Universal Robots URScript: FaiChun_9 Jan_11_2_t3.script

def Machining3():
  # Default parameters:
  global speed_ms = 0.05
  global speed_rads = 0.75
  global accel_mss = 3
  global accel_radss = 1.2
  global blend_radius_m = 0.0003

  # Add subprograms here
  # Start of main program
  # Program generated by RoboDK v5.6.8 for UR10e on 17/01/2025 15:25:47
  # Using nominal kinematics.
  blend_radius_m = 0.0003
  speed_ms = 0.05
  # set_reference(p[0.340000, 0.130000, 0.001500, 0.000000, 0.000000, 0.000000])
  set_tcp(p[0.000000, 0.000000, 0.252000, 0.000000, 0.000000, 0.000000])
  # Show Tool
  movej([0.835374, -1.505568, -2.356532, -0.850289, 1.570796, 2.406170],accel_radss,speed_rads,0,blend_radius_m)
  movel([0.835374, -1.553863, -2.383497, -0.775029, 1.570796, 2.406170],accel_mss,speed_ms,0,blend_radius_m)
  #SetTool1
  #M_RunCode6
  #SetRPM60000
  speed_ms = 0.05
  #M_RunCode3
  movel([0.835374, -1.574630, -2.393441, -0.744318, 1.570796, 2.406170],accel_mss,speed_ms,0,blend_radius_m)
  speed_ms = 0.003
  movel([0.835374, -1.579969, -2.395857, -0.736564, 1.570796, 2.406170],accel_mss,speed_ms,0,blend_radius_m)
  speed_ms = 0.015
  movel([0.633989, -1.489921, -2.480769, -0.741699, 1.570796, 2.204786],accel_mss,speed_ms,0,blend_radius_m)
  movel([0.864064, -1.190756, -2.677424, -0.844209, 1.570796, 2.434860],accel_mss,speed_ms,0,blend_radius_m)
  movel([1.072859, -1.363512, -2.578824, -0.770053, 1.570796, 2.643656],accel_mss,speed_ms,0,blend_radius_m)
  movel([0.835374, -1.579969, -2.395857, -0.736564, 1.570796, 2.406170],accel_mss,speed_ms,0,blend_radius_m)
  speed_ms = 0.003
  movel([0.835374, -1.574630, -2.393441, -0.744318, 1.570796, 2.406170],accel_mss,speed_ms,0,blend_radius_m)
  speed_ms = 0.05
  movel([0.835374, -1.553863, -2.383497, -0.775029, 1.570796, 2.406170],accel_mss,speed_ms,0,blend_radius_m)
  #M_RunCode9
  movel([0.837981, -1.545638, -2.391457, -0.775294, 1.570796, 2.408778],accel_mss,speed_ms,0,blend_radius_m)
  #M_RunCode3
  movel([0.837981, -1.566582, -2.401486, -0.744320, 1.570796, 2.408778],accel_mss,speed_ms,0,blend_radius_m)
  speed_ms = 0.003
  movel([0.837981, -1.571968, -2.403923, -0.736498, 1.570796, 2.408778],accel_mss,speed_ms,0,blend_radius_m)
  speed_ms = 0.012
  movel([0.835363, -1.570327, -2.405565, -0.736497, 1.570796, 2.406160],accel_mss,speed_ms,0,blend_radius_m)
  movel([0.832471, -1.573305, -2.402582, -0.736502, 1.570796, 2.403268],accel_mss,speed_ms,0,blend_radius_m)
  movel([0.828572, -1.570903, -2.404989, -0.736497, 1.570796, 2.399369],accel_mss,speed_ms,0,blend_radius_m)
  movel([0.831462, -1.567905, -2.407980, -0.736503, 1.570796, 2.402259],accel_mss,speed_ms,0,blend_radius_m)
  movel([0.830089, -1.567061, -2.408820, -0.736508, 1.570796, 2.400885],accel_mss,speed_ms,0,blend_radius_m)
  movel([0.827198, -1.570064, -2.405828, -0.736497, 1.570796, 2.397994],accel_mss,speed_ms,0,blend_radius_m)
  movel([0.823900, -1.568068, -2.407819, -0.736503, 1.570796, 2.394696],accel_mss,speed_ms,0,blend_radius_m)
  movel([0.823259, -1.567680, -2.408205, -0.736504, 1.570796, 2.394055],accel_mss,speed_ms,0,blend_radius_m)
  movel([0.827542, -1.563207, -2.412639, -0.736543, 1.570796, 2.398338],accel_mss,speed_ms,0,blend_radius_m)
  movel([0.830207, -1.564832, -2.411032, -0.736525, 1.570796, 2.401003],accel_mss,speed_ms,0,blend_radius_m)
  movel([0.831719, -1.563265, -2.412582, -0.736542, 1.570796, 2.402516],accel_mss,speed_ms,0,blend_radius_m)
  movel([0.827666, -1.560790, -2.415022, -0.736577, 1.570796, 2.398462],accel_mss,speed_ms,0,blend_radius_m)
  movel([0.821871, -1.566850, -2.409030, -0.736509, 1.570796, 2.392667],accel_mss,speed_ms,0,blend_radius_m)
  movel([0.821225, -1.566466, -2.409411, -0.736512, 1.570796, 2.392022],accel_mss,speed_ms,0,blend_radius_m)
  speed_ms = 0.02
  movel([0.744589, -1.526264, -2.448047, -0.738078, 1.570796, 2.315386],accel_mss,speed_ms,0,blend_radius_m)
  movel([0.657367, -1.492537, -2.478483, -0.741369, 1.570796, 2.228164],accel_mss,speed_ms,0,blend_radius_m)
  speed_ms = 0.012
  movel([0.662664, -1.485271, -2.484806, -0.742313, 1.570796, 2.233460],accel_mss,speed_ms,0,blend_radius_m)
  movel([0.657451, -1.483595, -2.486252, -0.742542, 1.570796, 2.228247],accel_mss,speed_ms,0,blend_radius_m)
  movel([0.656073, -1.485492, -2.484614, -0.742283, 1.570796, 2.226869],accel_mss,speed_ms,0,blend_radius_m)
  movel([0.659505, -1.486587, -2.483666, -0.742136, 1.570796, 2.230302],accel_mss,speed_ms,0,blend_radius_m)
  movel([0.655595, -1.491963, -2.478985, -0.741441, 1.570796, 2.226392],accel_mss,speed_ms,0,blend_radius_m)
  movel([0.654774, -1.491702, -2.479213, -0.741473, 1.570796, 2.225570],accel_mss,speed_ms,0,blend_radius_m)
  movel([0.650526, -1.490368, -2.480379, -0.741642, 1.570796, 2.221322],accel_mss,speed_ms,0,blend_radius_m)
  movel([0.653148, -1.486728, -2.483544, -0.742117, 1.570796, 2.223944],accel_mss,speed_ms,0,blend_radius_m)
  movel([0.651362, -1.486169, -2.484029, -0.742192, 1.570796, 2.222158],accel_mss,speed_ms,0,blend_radius_m)
  movel([0.648743, -1.489815, -2.480861, -0.741713, 1.570796, 2.219539],accel_mss,speed_ms,0,blend_radius_m)
  movel([0.643637, -1.488255, -2.482219, -0.741915, 1.570796, 2.214433],accel_mss,speed_ms,0,blend_radius_m)
  movel([0.646242, -1.484596, -2.485388, -0.742404, 1.570796, 2.217038],accel_mss,speed_ms,0,blend_radius_m)
  movel([0.642766, -1.483550, -2.486291, -0.742548, 1.570796, 2.213562],accel_mss,speed_ms,0,blend_radius_m)
  movel([0.646649, -1.478084, -2.490978, -0.743327, 1.570796, 2.217445],accel_mss,speed_ms,0,blend_radius_m)
  movel([0.650136, -1.479145, -2.490072, -0.743172, 1.570796, 2.220932],accel_mss,speed_ms,0,blend_radius_m)
  movel([0.651513, -1.477225, -2.491711, -0.743453, 1.570796, 2.222309],accel_mss,speed_ms,0,blend_radius_m)
  movel([0.648022, -1.476157, -2.492620, -0.743612, 1.570796, 2.218819],accel_mss,speed_ms,0,blend_radius_m)
  movel([0.651321, -1.471538, -2.496531, -0.744320, 1.570796, 2.222117],accel_mss,speed_ms,0,blend_radius_m)
  movel([0.651968, -1.470637, -2.497290, -0.744462, 1.570796, 2.222765],accel_mss,speed_ms,0,blend_radius_m)
  movel([0.657153, -1.472242, -2.495937, -0.744210, 1.570796, 2.227950],accel_mss,speed_ms,0,blend_radius_m)
  movel([0.654471, -1.475959, -2.492788, -0.743642, 1.570796, 2.225267],accel_mss,speed_ms,0,blend_radius_m)
  movel([0.656278, -1.476523, -2.492308, -0.743557, 1.570796, 2.227074],accel_mss,speed_ms,0,blend_radius_m)
  movel([0.660366, -1.470877, -2.497088, -0.744424, 1.570796, 2.231163],accel_mss,speed_ms,0,blend_radius_m)
  movel([0.653364, -1.468690, -2.498926, -0.744773, 1.570796, 2.224160],accel_mss,speed_ms,0,blend_radius_m)
  movel([0.735208, -1.358940, -2.581932, -0.771517, 1.570796, 2.306004],accel_mss,speed_ms,0,blend_radius_m)
  speed_ms = 0.02
  movel([0.838762, -1.228759, -2.658846, -0.824784, 1.570796, 2.409558],accel_mss,speed_ms,0,blend_radius_m)
  movel([0.839821, -1.227466, -2.659505, -0.825418, 1.570796, 2.410617],accel_mss,speed_ms,0,blend_radius_m)
  speed_ms = 0.012
  movel([0.847664, -1.231537, -2.657424, -0.823428, 1.570796, 2.418460],accel_mss,speed_ms,0,blend_radius_m)
  movel([0.854413, -1.223391, -2.661569, -0.827429, 1.570796, 2.425209],accel_mss,speed_ms,0,blend_radius_m)
  movel([0.852387, -1.222304, -2.662116, -0.827969, 1.570796, 2.423183],accel_mss,speed_ms,0,blend_radius_m)
  movel([0.847934, -1.227691, -2.659391, -0.825307, 1.570796, 2.418730],accel_mss,speed_ms,0,blend_radius_m)
  movel([0.842121, -1.224661, -2.660928, -0.826800, 1.570796, 2.412917],accel_mss,speed_ms,0,blend_radius_m)
  movel([0.843184, -1.223362, -2.661584, -0.827444, 1.570796, 2.413980],accel_mss,speed_ms,0,blend_radius_m)
  movel([0.848718, -1.216604, -2.664964, -0.830821, 1.570796, 2.419515],accel_mss,speed_ms,0,blend_radius_m)
  movel([0.852657, -1.218688, -2.663927, -0.829774, 1.570796, 2.423453],accel_mss,speed_ms,0,blend_radius_m)
  movel([0.854994, -1.215856, -2.665335, -0.831197, 1.570796, 2.425791],accel_mss,speed_ms,0,blend_radius_m)
  movel([0.851054, -1.213757, -2.666373, -0.832259, 1.570796, 2.421850],accel_mss,speed_ms,0,blend_radius_m)
  movel([0.857788, -1.205562, -2.670377, -0.836450, 1.570796, 2.428584],accel_mss,speed_ms,0,blend_radius_m)
  movel([0.861735, -1.207706, -2.669337, -0.835346, 1.570796, 2.432532],accel_mss,speed_ms,0,blend_radius_m)
  movel([0.866344, -1.202146, -2.672025, -0.838219, 1.570796, 2.437140],accel_mss,speed_ms,0,blend_radius_m)
  movel([0.872146, -1.205404, -2.670454, -0.836531, 1.570796, 2.442943],accel_mss,speed_ms,0,blend_radius_m)
  movel([0.867532, -1.210918, -2.667769, -0.833702, 1.570796, 2.438328],accel_mss,speed_ms,0,blend_radius_m)
  movel([0.869549, -1.212054, -2.667212, -0.833124, 1.570796, 2.440345],accel_mss,speed_ms,0,blend_radius_m)
  movel([0.874165, -1.206556, -2.669896, -0.835937, 1.570796, 2.444961],accel_mss,speed_ms,0,blend_radius_m)
  movel([0.879884, -1.209871, -2.668281, -0.834237, 1.570796, 2.450680],accel_mss,speed_ms,0,blend_radius_m)
  movel([0.873058, -1.217928, -2.664306, -0.830155, 1.570796, 2.443854],accel_mss,speed_ms,0,blend_radius_m)
  movel([0.869206, -1.215731, -2.665397, -0.831261, 1.570796, 2.440003],accel_mss,speed_ms,0,blend_radius_m)
  movel([0.866837, -1.218550, -2.663996, -0.829843, 1.570796, 2.437634],accel_mss,speed_ms,0,blend_radius_m)
  movel([0.872676, -1.221871, -2.662334, -0.828184, 1.570796, 2.443472],accel_mss,speed_ms,0,blend_radius_m)
  movel([0.881873, -1.211042, -2.667708, -0.833639, 1.570796, 2.452670],accel_mss,speed_ms,0,blend_radius_m)
  movel([0.975719, -1.277693, -2.632456, -0.802240, 1.570796, 2.546515],accel_mss,speed_ms,0,blend_radius_m)
  speed_ms = 0.02
  movel([1.052001, -1.350806, -2.587390, -0.774193, 1.570796, 2.622798],accel_mss,speed_ms,0,blend_radius_m)
  movel([1.043190, -1.358370, -2.582317, -0.771702, 1.570796, 2.613987],accel_mss,speed_ms,0,blend_radius_m)
  speed_ms = 0.012
  movel([1.047039, -1.362473, -2.579533, -0.770383, 1.570796, 2.617836],accel_mss,speed_ms,0,blend_radius_m)
  movel([1.049307, -1.360540, -2.580848, -0.771002, 1.570796, 2.620103],accel_mss,speed_ms,0,blend_radius_m)
  movel([1.046783, -1.357825, -2.582685, -0.771878, 1.570796, 2.617579],accel_mss,speed_ms,0,blend_radius_m)
  movel([1.053311, -1.352246, -2.586430, -0.773713, 1.570796, 2.624108],accel_mss,speed_ms,0,blend_radius_m)
  movel([1.053918, -1.352909, -2.585988, -0.773493, 1.570796, 2.624714],accel_mss,speed_ms,0,blend_radius_m)
  movel([1.057025, -1.356325, -2.583697, -0.772367, 1.570796, 2.627821],accel_mss,speed_ms,0,blend_radius_m)
  movel([1.052623, -1.360057, -2.581176, -0.771157, 1.570796, 2.623420],accel_mss,speed_ms,0,blend_radius_m)
  movel([1.053917, -1.361475, -2.580212, -0.770702, 1.570796, 2.624713],accel_mss,speed_ms,0,blend_radius_m)
  movel([1.058318, -1.357758, -2.582731, -0.771900, 1.570796, 2.629115],accel_mss,speed_ms,0,blend_radius_m)
  movel([1.061975, -1.361842, -2.579962, -0.770584, 1.570796, 2.632771],accel_mss,speed_ms,0,blend_radius_m)
  movel([1.057587, -1.365521, -2.577449, -0.769419, 1.570796, 2.628383],accel_mss,speed_ms,0,blend_radius_m)
  movel([1.060041, -1.368254, -2.575569, -0.768566, 1.570796, 2.630837],accel_mss,speed_ms,0,blend_radius_m)
  movel([1.053613, -1.373635, -2.571837, -0.766917, 1.570796, 2.624409],accel_mss,speed_ms,0,blend_radius_m)
  movel([1.051147, -1.370941, -2.573711, -0.767737, 1.570796, 2.621943],accel_mss,speed_ms,0,blend_radius_m)
  movel([1.048905, -1.372833, -2.572396, -0.767160, 1.570796, 2.619702],accel_mss,speed_ms,0,blend_radius_m)
  movel([1.051373, -1.375516, -2.570523, -0.766350, 1.570796, 2.622169],accel_mss,speed_ms,0,blend_radius_m)
  movel([1.046058, -1.379991, -2.567376, -0.765022, 1.570796, 2.616855],accel_mss,speed_ms,0,blend_radius_m)
  movel([1.045032, -1.380857, -2.566764, -0.764768, 1.570796, 2.615828],accel_mss,speed_ms,0,blend_radius_m)
  movel([1.041351, -1.376942, -2.569524, -0.765924, 1.570796, 2.612147],accel_mss,speed_ms,0,blend_radius_m)
  movel([1.045637, -1.373301, -2.572070, -0.767018, 1.570796, 2.616433],accel_mss,speed_ms,0,blend_radius_m)
  movel([1.044340, -1.371916, -2.573034, -0.767439, 1.570796, 2.615136],accel_mss,speed_ms,0,blend_radius_m)
  movel([1.037833, -1.377462, -2.569158, -0.765769, 1.570796, 2.608629],accel_mss,speed_ms,0,blend_radius_m)
  movel([1.042823, -1.382724, -2.565440, -0.764225, 1.570796, 2.613619],accel_mss,speed_ms,0,blend_radius_m)
  speed_ms = 0.02
  movel([0.937722, -1.475331, -2.493322, -0.743736, 1.570796, 2.508518],accel_mss,speed_ms,0,blend_radius_m)
  movel([0.849748, -1.560014, -2.415785, -0.736589, 1.570796, 2.420545],accel_mss,speed_ms,0,blend_radius_m)
  speed_ms = 0.012
  movel([0.844480, -1.556645, -2.419087, -0.736656, 1.570796, 2.415277],accel_mss,speed_ms,0,blend_radius_m)
  movel([0.839983, -1.561236, -2.414583, -0.736570, 1.570796, 2.410779],accel_mss,speed_ms,0,blend_radius_m)
  movel([0.841353, -1.562100, -2.413732, -0.736557, 1.570796, 2.412149],accel_mss,speed_ms,0,blend_radius_m)
  movel([0.844308, -1.559087, -2.416696, -0.736606, 1.570796, 2.415104],accel_mss,speed_ms,0,blend_radius_m)
  movel([0.848197, -1.561574, -2.414251, -0.736565, 1.570796, 2.418993],accel_mss,speed_ms,0,blend_radius_m)
  movel([0.847483, -1.562295, -2.413539, -0.736554, 1.570796, 2.418279],accel_mss,speed_ms,0,blend_radius_m)
  movel([0.843823, -1.566008, -2.409866, -0.736515, 1.570796, 2.414620],accel_mss,speed_ms,0,blend_radius_m)
  movel([0.841203, -1.564344, -2.411515, -0.736530, 1.570796, 2.411999],accel_mss,speed_ms,0,blend_radius_m)
  movel([0.839681, -1.565899, -2.409974, -0.736516, 1.570796, 2.410477],accel_mss,speed_ms,0,blend_radius_m)
  movel([0.842302, -1.567558, -2.408326, -0.736505, 1.570796, 2.413098],accel_mss,speed_ms,0,blend_radius_m)
  movel([0.837981, -1.571968, -2.403923, -0.736498, 1.570796, 2.408778],accel_mss,speed_ms,0,blend_radius_m)
  speed_ms = 0.003
  movel([0.837981, -1.566582, -2.401486, -0.744320, 1.570796, 2.408778],accel_mss,speed_ms,0,blend_radius_m)
  speed_ms = 0.05
  movel([0.837981, -1.545638, -2.391457, -0.775294, 1.570796, 2.408778],accel_mss,speed_ms,0,blend_radius_m)
  #M_RunCode9
  movel([0.855198, -1.260338, -2.606468, -0.845583, 1.570796, 2.425994],accel_mss,speed_ms,0,blend_radius_m)
  #M_RunCode3
  # num 0 inside
  movel([0.855198, -1.286686, -2.619958, -0.805745, 1.570796, 2.425994],accel_mss,speed_ms,0,blend_radius_m)
  speed_ms = 0.003
  movel([0.855198, -1.293571, -2.623261, -0.795557, 1.570796, 2.425994],accel_mss,speed_ms,0,blend_radius_m)
  speed_ms = 0.015
  movel([0.846910, -1.296288, -2.621656, -0.794445, 1.570796, 2.417706],accel_mss,speed_ms,0,blend_radius_m)
  movel([0.841111, -1.297727, -2.620801, -0.793860, 1.570796, 2.411907],accel_mss,speed_ms,0,blend_radius_m)
  movel([0.839123, -1.297920, -2.620687, -0.793782, 1.570796, 2.409919],accel_mss,speed_ms,0,blend_radius_m)
  movel([0.837725, -1.297694, -2.620821, -0.793874, 1.570796, 2.408522],accel_mss,speed_ms,0,blend_radius_m)
  movel([0.836916, -1.297054, -2.621202, -0.794134, 1.570796, 2.407712],accel_mss,speed_ms,0,blend_radius_m)
  movel([0.836696, -1.295992, -2.621831, -0.794566, 1.570796, 2.407493],accel_mss,speed_ms,0,blend_radius_m)
  movel([0.837055, -1.294718, -2.622585, -0.795086, 1.570796, 2.407851],accel_mss,speed_ms,0,blend_radius_m)
  movel([0.837982, -1.293440, -2.623338, -0.795611, 1.570796, 2.408779],accel_mss,speed_ms,0,blend_radius_m)
  movel([0.839480, -1.292159, -2.624092, -0.796138, 1.570796, 2.410276],accel_mss,speed_ms,0,blend_radius_m)
  movel([0.841550, -1.290874, -2.624846, -0.796670, 1.570796, 2.412346],accel_mss,speed_ms,0,blend_radius_m)
  movel([0.847491, -1.288081, -2.626476, -0.797832, 1.570796, 2.418287],accel_mss,speed_ms,0,blend_radius_m)
  movel([0.855893, -1.284860, -2.628345, -0.799184, 1.570796, 2.426689],accel_mss,speed_ms,0,blend_radius_m)
  movel([0.864286, -1.282119, -2.629925, -0.800345, 1.570796, 2.435082],accel_mss,speed_ms,0,blend_radius_m)
  movel([0.870165, -1.280730, -2.630722, -0.800937, 1.570796, 2.440961],accel_mss,speed_ms,0,blend_radius_m)
  movel([0.872167, -1.280581, -2.630807, -0.801001, 1.570796, 2.442964],accel_mss,speed_ms,0,blend_radius_m)
  movel([0.873560, -1.280853, -2.630651, -0.800885, 1.570796, 2.444356],accel_mss,speed_ms,0,blend_radius_m)
  movel([0.874341, -1.281545, -2.630255, -0.800590, 1.570796, 2.445137],accel_mss,speed_ms,0,blend_radius_m)
  movel([0.874513, -1.282655, -2.629617, -0.800118, 1.570796, 2.445309],accel_mss,speed_ms,0,blend_radius_m)
  movel([0.874099, -1.283962, -2.628863, -0.799563, 1.570796, 2.444895],accel_mss,speed_ms,0,blend_radius_m)
  movel([0.873124, -1.285249, -2.628120, -0.799020, 1.570796, 2.443921],accel_mss,speed_ms,0,blend_radius_m)
  movel([0.871587, -1.286518, -2.627385, -0.798486, 1.570796, 2.442383],accel_mss,speed_ms,0,blend_radius_m)
  movel([0.869494, -1.287766, -2.626660, -0.797963, 1.570796, 2.440290],accel_mss,speed_ms,0,blend_radius_m)
  movel([0.863543, -1.290454, -2.625092, -0.796844, 1.570796, 2.434339],accel_mss,speed_ms,0,blend_radius_m)
  movel([0.855198, -1.293571, -2.623261, -0.795557, 1.570796, 2.425994],accel_mss,speed_ms,0,blend_radius_m)
  speed_ms = 0.003
  movel([0.855198, -1.286686, -2.619958, -0.805745, 1.570796, 2.425994],accel_mss,speed_ms,0,blend_radius_m)
  speed_ms = 0.05
  movel([0.855198, -1.260338, -2.606468, -0.845583, 1.570796, 2.425994],accel_mss,speed_ms,0,blend_radius_m)
  #M_RunCode9
  movel([0.854459, -1.269799, -2.601095, -0.841495, 1.570796, 2.425256],accel_mss,speed_ms,0,blend_radius_m)
  #M_RunCode3
  #num 0 outside
  movel([0.854459, -1.296016, -2.614460, -0.801913, 1.570796, 2.425256],accel_mss,speed_ms,0,blend_radius_m)
  speed_ms = 0.003
  movel([0.854459, -1.302862, -2.617732, -0.791795, 1.570796, 2.425256],accel_mss,speed_ms,0,blend_radius_m)
  speed_ms = 0.015
  movel([0.851475, -1.303789, -2.617174, -0.791426, 1.570796, 2.422272],accel_mss,speed_ms,0,blend_radius_m)
  movel([0.848730, -1.304421, -2.616793, -0.791175, 1.570796, 2.419526],accel_mss,speed_ms,0,blend_radius_m)
  movel([0.846217, -1.304761, -2.616588, -0.791040, 1.570796, 2.417014],accel_mss,speed_ms,0,blend_radius_m)
  movel([0.843939, -1.304807, -2.616560, -0.791022, 1.570796, 2.414735],accel_mss,speed_ms,0,blend_radius_m)
  movel([0.841916, -1.304581, -2.616697, -0.791111, 1.570796, 2.412713],accel_mss,speed_ms,0,blend_radius_m)
  movel([0.840172, -1.304105, -2.616984, -0.791300, 1.570796, 2.410968],accel_mss,speed_ms,0,blend_radius_m)
  movel([0.838702, -1.303380, -2.617420, -0.791589, 1.570796, 2.409498],accel_mss,speed_ms,0,blend_radius_m)
  movel([0.837514, -1.302400, -2.618010, -0.791979, 1.570796, 2.408310],accel_mss,speed_ms,0,blend_radius_m)
  movel([0.836610, -1.301192, -2.618734, -0.792463, 1.570796, 2.407406],accel_mss,speed_ms,0,blend_radius_m)
  movel([0.835994, -1.299790, -2.619572, -0.793026, 1.570796, 2.406790],accel_mss,speed_ms,0,blend_radius_m)
  movel([0.835668, -1.298186, -2.620529, -0.793674, 1.570796, 2.406464],accel_mss,speed_ms,0,blend_radius_m)
  movel([0.835631, -1.296383, -2.621599, -0.794407, 1.570796, 2.406427],accel_mss,speed_ms,0,blend_radius_m)
  movel([0.835884, -1.294466, -2.622733, -0.795190, 1.570796, 2.406680],accel_mss,speed_ms,0,blend_radius_m)
  movel([0.836421, -1.292534, -2.623871, -0.795983, 1.570796, 2.407217],accel_mss,speed_ms,0,blend_radius_m)
  movel([0.837240, -1.290586, -2.625014, -0.796789, 1.570796, 2.408036],accel_mss,speed_ms,0,blend_radius_m)
  movel([0.838350, -1.288617, -2.626164, -0.797608, 1.570796, 2.409146],accel_mss,speed_ms,0,blend_radius_m)
  movel([0.839739, -1.286668, -2.627298, -0.798423, 1.570796, 2.410536],accel_mss,speed_ms,0,blend_radius_m)
  movel([0.841401, -1.284772, -2.628396, -0.799221, 1.570796, 2.412197],accel_mss,speed_ms,0,blend_radius_m)
  movel([0.843338, -1.282931, -2.629458, -0.800000, 1.570796, 2.414134],accel_mss,speed_ms,0,blend_radius_m)
  movel([0.845550, -1.281147, -2.630483, -0.800759, 1.570796, 2.416347],accel_mss,speed_ms,0,blend_radius_m)
  movel([0.848009, -1.279462, -2.631447, -0.801480, 1.570796, 2.418805],accel_mss,speed_ms,0,blend_radius_m)
  movel([0.850682, -1.277926, -2.632323, -0.802140, 1.570796, 2.421478],accel_mss,speed_ms,0,blend_radius_m)
  movel([0.853567, -1.276542, -2.633110, -0.802737, 1.570796, 2.424364],accel_mss,speed_ms,0,blend_radius_m)
  movel([0.856663, -1.275312, -2.633807, -0.803270, 1.570796, 2.427459],accel_mss,speed_ms,0,blend_radius_m)
  movel([0.859747, -1.274318, -2.634369, -0.803702, 1.570796, 2.430544],accel_mss,speed_ms,0,blend_radius_m)
  movel([0.862585, -1.273645, -2.634749, -0.803995, 1.570796, 2.433381],accel_mss,speed_ms,0,blend_radius_m)
  movel([0.865178, -1.273292, -2.634948, -0.804149, 1.570796, 2.435974],accel_mss,speed_ms,0,blend_radius_m)
  movel([0.867519, -1.273260, -2.634966, -0.804163, 1.570796, 2.438315],accel_mss,speed_ms,0,blend_radius_m)
  movel([0.869584, -1.273524, -2.634817, -0.804048, 1.570796, 2.440380],accel_mss,speed_ms,0,blend_radius_m)
  movel([0.871341, -1.274060, -2.634515, -0.803814, 1.570796, 2.442138],accel_mss,speed_ms,0,blend_radius_m)
  movel([0.872797, -1.274863, -2.634061, -0.803465, 1.570796, 2.443593],accel_mss,speed_ms,0,blend_radius_m)
  movel([0.873946, -1.275936, -2.633454, -0.803000, 1.570796, 2.444743],accel_mss,speed_ms,0,blend_radius_m)
  movel([0.874790, -1.277237, -2.632715, -0.802437, 1.570796, 2.445586],accel_mss,speed_ms,0,blend_radius_m)
  movel([0.875334, -1.278736, -2.631862, -0.801792, 1.570796, 2.446131],accel_mss,speed_ms,0,blend_radius_m)
  movel([0.875580, -1.280428, -2.630895, -0.801066, 1.570796, 2.446377],accel_mss,speed_ms,0,blend_radius_m)
  movel([0.875527, -1.282310, -2.629815, -0.800264, 1.570796, 2.446323],accel_mss,speed_ms,0,blend_radius_m)
  movel([0.875187, -1.284285, -2.628677, -0.799427, 1.570796, 2.445983],accel_mss,speed_ms,0,blend_radius_m)
  movel([0.874574, -1.286253, -2.627538, -0.798598, 1.570796, 2.445370],accel_mss,speed_ms,0,blend_radius_m)
  movel([0.873688, -1.288215, -2.626398, -0.797776, 1.570796, 2.444484],accel_mss,speed_ms,0,blend_radius_m)
  movel([0.872531, -1.290171, -2.625257, -0.796961, 1.570796, 2.443327],accel_mss,speed_ms,0,blend_radius_m)
  movel([0.871111, -1.292085, -2.624135, -0.796169, 1.570796, 2.441907],accel_mss,speed_ms,0,blend_radius_m)
  movel([0.869432, -1.293928, -2.623051, -0.795410, 1.570796, 2.440228],accel_mss,speed_ms,0,blend_radius_m)
  movel([0.867493, -1.295700, -2.622004, -0.794685, 1.570796, 2.438289],accel_mss,speed_ms,0,blend_radius_m)
  movel([0.865298, -1.297400, -2.620996, -0.793993, 1.570796, 2.436095],accel_mss,speed_ms,0,blend_radius_m)
  movel([0.862881, -1.298989, -2.620050, -0.793350, 1.570796, 2.433677],accel_mss,speed_ms,0,blend_radius_m)
  movel([0.860267, -1.300428, -2.619191, -0.792770, 1.570796, 2.431063],accel_mss,speed_ms,0,blend_radius_m)
  movel([0.857460, -1.301718, -2.618419, -0.792252, 1.570796, 2.428257],accel_mss,speed_ms,0,blend_radius_m)
  movel([0.854459, -1.302862, -2.617732, -0.791795, 1.570796, 2.425256],accel_mss,speed_ms,0,blend_radius_m)
  speed_ms = 0.003
  movel([0.854459, -1.296016, -2.614460, -0.801913, 1.570796, 2.425256],accel_mss,speed_ms,0,blend_radius_m)
  speed_ms = 0.05
  movel([0.854459, -1.269799, -2.601095, -0.841495, 1.570796, 2.425256],accel_mss,speed_ms,0,blend_radius_m)
  #M_RunCode9
  movel([0.848212, -1.241330, -2.616943, -0.854116, 1.570796, 2.419008],accel_mss,speed_ms,0,blend_radius_m)
  #M_RunCode3
  # num 2
  movel([0.848212, -1.267925, -2.630682, -0.813782, 1.570796, 2.419008],accel_mss,speed_ms,0,blend_radius_m)
  speed_ms = 0.003
  movel([0.848212, -1.274884, -2.634049, -0.803455, 1.570796, 2.419008],accel_mss,speed_ms,0,blend_radius_m)
  speed_ms = 0.02
  movel([0.837317, -1.278925, -2.631754, -0.801710, 1.570796, 2.408113],accel_mss,speed_ms,0,blend_radius_m)
  movel([0.839074, -1.249773, -2.647865, -0.814751, 1.570796, 2.409870],accel_mss,speed_ms,0,blend_radius_m)
  movel([0.840196, -1.249335, -2.648099, -0.814955, 1.570796, 2.410992],accel_mss,speed_ms,0,blend_radius_m)
  movel([0.843034, -1.248564, -2.648511, -0.815314, 1.570796, 2.413831],accel_mss,speed_ms,0,blend_radius_m)
  movel([0.845771, -1.248506, -2.648542, -0.815341, 1.570796, 2.416567],accel_mss,speed_ms,0,blend_radius_m)
  movel([0.848339, -1.248990, -2.648284, -0.815116, 1.570796, 2.419136],accel_mss,speed_ms,0,blend_radius_m)
  movel([0.850670, -1.249839, -2.647829, -0.814720, 1.570796, 2.421467],accel_mss,speed_ms,0,blend_radius_m)
  movel([0.856325, -1.252900, -2.646186, -0.813303, 1.570796, 2.427121],accel_mss,speed_ms,0,blend_radius_m)
  movel([0.861461, -1.255841, -2.644597, -0.811951, 1.570796, 2.432257],accel_mss,speed_ms,0,blend_radius_m)
  movel([0.863580, -1.256692, -2.644135, -0.811562, 1.570796, 2.434377],accel_mss,speed_ms,0,blend_radius_m)
  movel([0.865859, -1.257203, -2.643857, -0.811329, 1.570796, 2.436655],accel_mss,speed_ms,0,blend_radius_m)
  movel([0.868233, -1.257243, -2.643835, -0.811311, 1.570796, 2.439030],accel_mss,speed_ms,0,blend_radius_m)
  movel([0.870648, -1.256675, -2.644144, -0.811570, 1.570796, 2.441444],accel_mss,speed_ms,0,blend_radius_m)
  movel([0.873569, -1.255238, -2.644923, -0.812228, 1.570796, 2.444365],accel_mss,speed_ms,0,blend_radius_m)
  movel([0.874767, -1.254321, -2.645420, -0.812649, 1.570796, 2.445563],accel_mss,speed_ms,0,blend_radius_m)
  movel([0.875791, -1.253271, -2.645986, -0.813132, 1.570796, 2.446587],accel_mss,speed_ms,0,blend_radius_m)
  movel([0.877258, -1.251040, -2.647186, -0.814163, 1.570796, 2.448054],accel_mss,speed_ms,0,blend_radius_m)
  movel([0.877898, -1.248826, -2.648371, -0.815192, 1.570796, 2.448694],accel_mss,speed_ms,0,blend_radius_m)
  movel([0.877875, -1.247491, -2.649083, -0.815815, 1.570796, 2.448671],accel_mss,speed_ms,0,blend_radius_m)
  movel([0.877482, -1.246635, -2.649538, -0.816216, 1.570796, 2.448278],accel_mss,speed_ms,0,blend_radius_m)
  movel([0.876798, -1.246264, -2.649735, -0.816390, 1.570796, 2.447594],accel_mss,speed_ms,0,blend_radius_m)
  movel([0.875913, -1.246377, -2.649675, -0.816337, 1.570796, 2.446709],accel_mss,speed_ms,0,blend_radius_m)
  movel([0.874526, -1.247366, -2.649149, -0.815874, 1.570796, 2.445322],accel_mss,speed_ms,0,blend_radius_m)
  movel([0.873202, -1.248420, -2.648588, -0.815381, 1.570796, 2.443999],accel_mss,speed_ms,0,blend_radius_m)
  movel([0.871495, -1.249252, -2.648143, -0.814993, 1.570796, 2.442292],accel_mss,speed_ms,0,blend_radius_m)
  movel([0.869538, -1.249620, -2.647947, -0.814822, 1.570796, 2.440334],accel_mss,speed_ms,0,blend_radius_m)
  movel([0.868153, -1.249104, -2.648222, -0.815062, 1.570796, 2.438950],accel_mss,speed_ms,0,blend_radius_m)
  movel([0.867374, -1.247895, -2.648867, -0.815626, 1.570796, 2.438171],accel_mss,speed_ms,0,blend_radius_m)
  movel([0.867234, -1.246189, -2.649775, -0.816425, 1.570796, 2.438030],accel_mss,speed_ms,0,blend_radius_m)
  movel([0.867710, -1.244254, -2.650799, -0.817336, 1.570796, 2.438506],accel_mss,speed_ms,0,blend_radius_m)
  movel([0.868781, -1.242353, -2.651802, -0.818234, 1.570796, 2.439578],accel_mss,speed_ms,0,blend_radius_m)
  movel([0.870379, -1.240727, -2.652656, -0.819006, 1.570796, 2.441175],accel_mss,speed_ms,0,blend_radius_m)
  movel([0.872426, -1.239628, -2.653231, -0.819530, 1.570796, 2.443223],accel_mss,speed_ms,0,blend_radius_m)
  movel([0.874179, -1.239185, -2.653463, -0.819741, 1.570796, 2.444975],accel_mss,speed_ms,0,blend_radius_m)
  movel([0.875671, -1.239239, -2.653435, -0.819716, 1.570796, 2.446467],accel_mss,speed_ms,0,blend_radius_m)
  movel([0.876905, -1.239788, -2.653148, -0.819454, 1.570796, 2.447701],accel_mss,speed_ms,0,blend_radius_m)
  movel([0.877875, -1.240835, -2.652599, -0.818955, 1.570796, 2.448672],accel_mss,speed_ms,0,blend_radius_m)
  movel([0.878573, -1.242283, -2.651839, -0.818268, 1.570796, 2.449370],accel_mss,speed_ms,0,blend_radius_m)
  movel([0.878998, -1.244031, -2.650917, -0.817441, 1.570796, 2.449794],accel_mss,speed_ms,0,blend_radius_m)
  movel([0.879021, -1.248427, -2.648584, -0.815378, 1.570796, 2.449817],accel_mss,speed_ms,0,blend_radius_m)
  movel([0.878543, -1.251428, -2.646978, -0.813983, 1.570796, 2.449340],accel_mss,speed_ms,0,blend_radius_m)
  movel([0.877746, -1.254377, -2.645389, -0.812623, 1.570796, 2.448542],accel_mss,speed_ms,0,blend_radius_m)
  movel([0.876632, -1.257271, -2.643820, -0.811298, 1.570796, 2.447428],accel_mss,speed_ms,0,blend_radius_m)
  movel([0.875201, -1.260113, -2.642269, -0.810007, 1.570796, 2.445997],accel_mss,speed_ms,0,blend_radius_m)
  movel([0.873417, -1.262713, -2.640842, -0.808835, 1.570796, 2.444214],accel_mss,speed_ms,0,blend_radius_m)
  movel([0.871230, -1.264887, -2.639642, -0.807860, 1.570796, 2.442027],accel_mss,speed_ms,0,blend_radius_m)
  movel([0.868642, -1.266641, -2.638669, -0.807078, 1.570796, 2.439438],accel_mss,speed_ms,0,blend_radius_m)
  movel([0.865652, -1.267984, -2.637922, -0.806483, 1.570796, 2.436448],accel_mss,speed_ms,0,blend_radius_m)
  movel([0.862952, -1.268698, -2.637524, -0.806167, 1.570796, 2.433748],accel_mss,speed_ms,0,blend_radius_m)
  movel([0.860488, -1.268833, -2.637449, -0.806107, 1.570796, 2.431284],accel_mss,speed_ms,0,blend_radius_m)
  movel([0.858259, -1.268518, -2.637624, -0.806246, 1.570796, 2.429055],accel_mss,speed_ms,0,blend_radius_m)
  movel([0.856267, -1.267886, -2.637977, -0.806526, 1.570796, 2.427063],accel_mss,speed_ms,0,blend_radius_m)
  movel([0.851897, -1.265592, -2.639251, -0.807546, 1.570796, 2.422694],accel_mss,speed_ms,0,blend_radius_m)
  movel([0.847719, -1.263475, -2.640421, -0.808492, 1.570796, 2.418515],accel_mss,speed_ms,0,blend_radius_m)
  movel([0.845888, -1.262909, -2.640734, -0.808746, 1.570796, 2.416685],accel_mss,speed_ms,0,blend_radius_m)
  movel([0.843868, -1.262640, -2.640882, -0.808867, 1.570796, 2.414664],accel_mss,speed_ms,0,blend_radius_m)
  movel([0.841671, -1.262784, -2.640803, -0.808803, 1.570796, 2.412467],accel_mss,speed_ms,0,blend_radius_m)
  movel([0.839325, -1.263447, -2.640437, -0.808505, 1.570796, 2.410122],accel_mss,speed_ms,0,blend_radius_m)
  movel([0.839258, -1.264541, -2.639833, -0.808015, 1.570796, 2.410054],accel_mss,speed_ms,0,blend_radius_m)
  movel([0.839240, -1.267497, -2.638194, -0.806699, 1.570796, 2.410037],accel_mss,speed_ms,0,blend_radius_m)
  movel([0.839588, -1.269943, -2.636829, -0.805617, 1.570796, 2.410384],accel_mss,speed_ms,0,blend_radius_m)
  movel([0.840292, -1.271889, -2.635738, -0.804762, 1.570796, 2.411089],accel_mss,speed_ms,0,blend_radius_m)
  movel([0.841357, -1.273337, -2.634923, -0.804129, 1.570796, 2.412154],accel_mss,speed_ms,0,blend_radius_m)
  movel([0.842716, -1.274334, -2.634360, -0.803695, 1.570796, 2.413512],accel_mss,speed_ms,0,blend_radius_m)
  movel([0.844310, -1.274923, -2.634027, -0.803439, 1.570796, 2.415107],accel_mss,speed_ms,0,blend_radius_m)
  movel([0.846140, -1.275106, -2.633924, -0.803359, 1.570796, 2.416937],accel_mss,speed_ms,0,blend_radius_m)
  movel([0.848212, -1.274884, -2.634049, -0.803455, 1.570796, 2.419008],accel_mss,speed_ms,0,blend_radius_m)
  speed_ms = 0.003
  movel([0.848212, -1.267925, -2.630682, -0.813782, 1.570796, 2.419008],accel_mss,speed_ms,0,blend_radius_m)
  speed_ms = 0.05
  movel([0.848212, -1.241330, -2.616943, -0.854116, 1.570796, 2.419008],accel_mss,speed_ms,0,blend_radius_m)
  #M_RunCode9
  movel([0.826211, -1.482495, -2.449132, -0.780763, 1.570796, 2.397007],accel_mss,speed_ms,0,blend_radius_m)
  #M_RunCode3
  movel([0.826211, -1.504789, -2.459853, -0.747747, 1.570796, 2.397007],accel_mss,speed_ms,0,blend_radius_m)
  speed_ms = 0.003
  movel([0.826211, -1.510538, -2.462462, -0.739389, 1.570796, 2.397007],accel_mss,speed_ms,0,blend_radius_m)
  speed_ms = 0.02
  movel([0.828289, -1.510208, -2.462760, -0.739421, 1.570796, 2.399085],accel_mss,speed_ms,0,blend_radius_m)
  movel([0.830302, -1.510363, -2.462620, -0.739406, 1.570796, 2.401099],accel_mss,speed_ms,0,blend_radius_m)
  movel([0.832201, -1.510879, -2.462153, -0.739357, 1.570796, 2.402998],accel_mss,speed_ms,0,blend_radius_m)
  movel([0.833928, -1.511634, -2.461469, -0.739285, 1.570796, 2.404725],accel_mss,speed_ms,0,blend_radius_m)
  movel([0.838141, -1.514151, -2.459185, -0.739053, 1.570796, 2.408937],accel_mss,speed_ms,0,blend_radius_m)
  movel([0.841979, -1.516541, -2.457006, -0.738842, 1.570796, 2.412776],accel_mss,speed_ms,0,blend_radius_m)
  movel([0.843557, -1.517276, -2.456333, -0.738779, 1.570796, 2.414353],accel_mss,speed_ms,0,blend_radius_m)
  movel([0.845249, -1.517784, -2.455869, -0.738736, 1.570796, 2.416045],accel_mss,speed_ms,0,blend_radius_m)
  movel([0.847003, -1.517969, -2.455699, -0.738721, 1.570796, 2.417800],accel_mss,speed_ms,0,blend_radius_m)
  movel([0.848777, -1.517734, -2.455914, -0.738741, 1.570796, 2.419573],accel_mss,speed_ms,0,blend_radius_m)
  movel([0.850907, -1.516929, -2.456651, -0.738809, 1.570796, 2.421703],accel_mss,speed_ms,0,blend_radius_m)
  movel([0.851774, -1.516373, -2.457159, -0.738857, 1.570796, 2.422570],accel_mss,speed_ms,0,blend_radius_m)
  movel([0.852509, -1.515713, -2.457761, -0.738914, 1.570796, 2.423305],accel_mss,speed_ms,0,blend_radius_m)
  movel([0.853547, -1.514267, -2.459079, -0.739043, 1.570796, 2.424343],accel_mss,speed_ms,0,blend_radius_m)
  movel([0.853974, -1.512781, -2.460429, -0.739178, 1.570796, 2.424770],accel_mss,speed_ms,0,blend_radius_m)
  movel([0.853932, -1.511858, -2.461267, -0.739264, 1.570796, 2.424728],accel_mss,speed_ms,0,blend_radius_m)
  movel([0.853622, -1.511243, -2.461824, -0.739322, 1.570796, 2.424418],accel_mss,speed_ms,0,blend_radius_m)
  movel([0.853113, -1.510942, -2.462096, -0.739351, 1.570796, 2.423910],accel_mss,speed_ms,0,blend_radius_m)
  movel([0.852463, -1.510961, -2.462079, -0.739349, 1.570796, 2.423260],accel_mss,speed_ms,0,blend_radius_m)
  movel([0.851461, -1.511551, -2.461545, -0.739293, 1.570796, 2.422258],accel_mss,speed_ms,0,blend_radius_m)
  movel([0.850505, -1.512192, -2.460964, -0.739233, 1.570796, 2.421301],accel_mss,speed_ms,0,blend_radius_m)
  movel([0.849263, -1.512650, -2.460549, -0.739190, 1.570796, 2.420059],accel_mss,speed_ms,0,blend_radius_m)
  movel([0.847827, -1.512776, -2.460434, -0.739179, 1.570796, 2.418623],accel_mss,speed_ms,0,blend_radius_m)
  movel([0.846798, -1.512325, -2.460843, -0.739221, 1.570796, 2.417595],accel_mss,speed_ms,0,blend_radius_m)
  movel([0.846201, -1.511436, -2.461649, -0.739304, 1.570796, 2.416998],accel_mss,speed_ms,0,blend_radius_m)
  movel([0.846067, -1.510252, -2.462720, -0.739417, 1.570796, 2.416863],accel_mss,speed_ms,0,blend_radius_m)
  movel([0.846384, -1.508949, -2.463897, -0.739544, 1.570796, 2.417180],accel_mss,speed_ms,0,blend_radius_m)
  movel([0.847138, -1.507712, -2.465010, -0.739666, 1.570796, 2.417934],accel_mss,speed_ms,0,blend_radius_m)
  movel([0.848281, -1.506704, -2.465916, -0.739768, 1.570796, 2.419077],accel_mss,speed_ms,0,blend_radius_m)
  movel([0.849765, -1.506089, -2.466469, -0.739831, 1.570796, 2.420561],accel_mss,speed_ms,0,blend_radius_m)
  movel([0.851044, -1.505901, -2.466638, -0.739851, 1.570796, 2.421841],accel_mss,speed_ms,0,blend_radius_m)
  movel([0.852144, -1.506039, -2.466514, -0.739836, 1.570796, 2.422940],accel_mss,speed_ms,0,blend_radius_m)
  movel([0.853060, -1.506500, -2.466100, -0.739789, 1.570796, 2.423856],accel_mss,speed_ms,0,blend_radius_m)
  movel([0.853793, -1.507282, -2.465397, -0.739710, 1.570796, 2.424590],accel_mss,speed_ms,0,blend_radius_m)
  movel([0.854338, -1.508321, -2.464463, -0.739606, 1.570796, 2.425134],accel_mss,speed_ms,0,blend_radius_m)
  movel([0.854685, -1.509551, -2.463353, -0.739485, 1.570796, 2.425481],accel_mss,speed_ms,0,blend_radius_m)
  movel([0.854795, -1.512578, -2.460614, -0.739197, 1.570796, 2.425591],accel_mss,speed_ms,0,blend_radius_m)
  movel([0.854503, -1.514619, -2.458759, -0.739011, 1.570796, 2.425299],accel_mss,speed_ms,0,blend_radius_m)
  movel([0.853974, -1.516606, -2.456946, -0.738837, 1.570796, 2.424771],accel_mss,speed_ms,0,blend_radius_m)
  movel([0.853209, -1.518538, -2.455178, -0.738673, 1.570796, 2.424006],accel_mss,speed_ms,0,blend_radius_m)
  movel([0.852208, -1.520418, -2.453452, -0.738520, 1.570796, 2.423004],accel_mss,speed_ms,0,blend_radius_m)
  movel([0.850938, -1.522109, -2.451894, -0.738386, 1.570796, 2.421734],accel_mss,speed_ms,0,blend_radius_m)
  movel([0.849360, -1.523482, -2.450625, -0.738281, 1.570796, 2.420156],accel_mss,speed_ms,0,blend_radius_m)
  movel([0.847476, -1.524539, -2.449647, -0.738203, 1.570796, 2.418273],accel_mss,speed_ms,0,blend_radius_m)
  movel([0.845283, -1.525282, -2.448959, -0.738148, 1.570796, 2.416080],accel_mss,speed_ms,0,blend_radius_m)
  movel([0.843296, -1.525606, -2.448658, -0.738125, 1.570796, 2.414093],accel_mss,speed_ms,0,blend_radius_m)
  movel([0.841472, -1.525538, -2.448721, -0.738130, 1.570796, 2.412269],accel_mss,speed_ms,0,blend_radius_m)
  movel([0.839814, -1.525169, -2.449063, -0.738156, 1.570796, 2.410611],accel_mss,speed_ms,0,blend_radius_m)
  movel([0.838330, -1.524594, -2.449596, -0.738198, 1.570796, 2.409126],accel_mss,speed_ms,0,blend_radius_m)
  movel([0.835060, -1.522694, -2.451354, -0.738341, 1.570796, 2.405857],accel_mss,speed_ms,0,blend_radius_m)
  movel([0.831940, -1.520927, -2.452983, -0.738479, 1.570796, 2.402736],accel_mss,speed_ms,0,blend_radius_m)
  movel([0.830580, -1.520402, -2.453466, -0.738521, 1.570796, 2.401376],accel_mss,speed_ms,0,blend_radius_m)
  movel([0.829081, -1.520075, -2.453766, -0.738547, 1.570796, 2.399877],accel_mss,speed_ms,0,blend_radius_m)
  movel([0.827459, -1.520022, -2.453815, -0.738551, 1.570796, 2.398255],accel_mss,speed_ms,0,blend_radius_m)
  movel([0.825733, -1.520322, -2.453539, -0.738527, 1.570796, 2.396530],accel_mss,speed_ms,0,blend_radius_m)
  movel([0.825695, -1.521083, -2.452839, -0.738467, 1.570796, 2.396491],accel_mss,speed_ms,0,blend_radius_m)
  movel([0.825719, -1.523155, -2.450928, -0.738306, 1.570796, 2.396516],accel_mss,speed_ms,0,blend_radius_m)
  movel([0.826004, -1.524901, -2.449312, -0.738176, 1.570796, 2.396800],accel_mss,speed_ms,0,blend_radius_m)
  movel([0.826548, -1.526318, -2.447997, -0.738074, 1.570796, 2.397345],accel_mss,speed_ms,0,blend_radius_m)
  movel([0.827354, -1.527411, -2.446980, -0.737997, 1.570796, 2.398150],accel_mss,speed_ms,0,blend_radius_m)
  movel([0.828375, -1.528207, -2.446239, -0.737943, 1.570796, 2.399171],accel_mss,speed_ms,0,blend_radius_m)
  movel([0.829564, -1.528731, -2.445750, -0.737908, 1.570796, 2.400360],accel_mss,speed_ms,0,blend_radius_m)
  movel([0.830926, -1.528985, -2.445514, -0.737891, 1.570796, 2.401722],accel_mss,speed_ms,0,blend_radius_m)
  movel([0.832458, -1.528968, -2.445530, -0.737892, 1.570796, 2.403255],accel_mss,speed_ms,0,blend_radius_m)
  movel([0.824422, -1.531079, -2.443555, -0.737755, 1.570796, 2.395218],accel_mss,speed_ms,0,blend_radius_m)
  movel([0.825388, -1.510763, -2.462259, -0.739368, 1.570796, 2.396184],accel_mss,speed_ms,0,blend_radius_m)
  movel([0.826211, -1.510538, -2.462462, -0.739389, 1.570796, 2.397007],accel_mss,speed_ms,0,blend_radius_m)
  speed_ms = 0.003
  movel([0.826211, -1.504789, -2.459853, -0.747747, 1.570796, 2.397007],accel_mss,speed_ms,0,blend_radius_m)
  speed_ms = 0.05
  movel([0.826211, -1.482495, -2.449132, -0.780763, 1.570796, 2.397007],accel_mss,speed_ms,0,blend_radius_m)
  #M_RunCode9
  movel([0.829309, -1.504822, -2.429429, -0.778138, 1.570796, 2.400105],accel_mss,speed_ms,0,blend_radius_m)
  #M_RunCode3
  movel([0.829309, -1.526641, -2.439900, -0.745848, 1.570796, 2.400105],accel_mss,speed_ms,0,blend_radius_m)
  speed_ms = 0.003
  movel([0.829309, -1.532262, -2.442446, -0.737681, 1.570796, 2.400105],accel_mss,speed_ms,0,blend_radius_m)
  speed_ms = 0.02
  movel([0.830725, -1.532125, -2.442575, -0.737689, 1.570796, 2.401522],accel_mss,speed_ms,0,blend_radius_m)
  movel([0.831763, -1.532549, -2.442177, -0.737663, 1.570796, 2.402559],accel_mss,speed_ms,0,blend_radius_m)
  movel([0.832382, -1.533401, -2.441376, -0.737612, 1.570796, 2.403178],accel_mss,speed_ms,0,blend_radius_m)
  movel([0.832538, -1.534548, -2.440297, -0.737545, 1.570796, 2.403335],accel_mss,speed_ms,0,blend_radius_m)
  movel([0.832247, -1.535806, -2.439110, -0.737473, 1.570796, 2.403043],accel_mss,speed_ms,0,blend_radius_m)
  movel([0.831515, -1.537002, -2.437979, -0.737408, 1.570796, 2.402312],accel_mss,speed_ms,0,blend_radius_m)
  movel([0.830408, -1.537979, -2.437054, -0.737356, 1.570796, 2.401204],accel_mss,speed_ms,0,blend_radius_m)
  movel([0.828978, -1.538578, -2.436486, -0.737325, 1.570796, 2.399775],accel_mss,speed_ms,0,blend_radius_m)
  movel([0.827793, -1.538742, -2.436331, -0.737316, 1.570796, 2.398589],accel_mss,speed_ms,0,blend_radius_m)
  movel([0.826918, -1.538583, -2.436482, -0.737324, 1.570796, 2.397714],accel_mss,speed_ms,0,blend_radius_m)
  movel([0.825989, -1.538499, -2.436561, -0.737329, 1.570796, 2.396785],accel_mss,speed_ms,0,blend_radius_m)
  movel([0.825341, -1.538812, -2.436265, -0.737313, 1.570796, 2.396138],accel_mss,speed_ms,0,blend_radius_m)
  movel([0.824793, -1.539384, -2.435721, -0.737284, 1.570796, 2.395589],accel_mss,speed_ms,0,blend_radius_m)
  movel([0.824409, -1.540106, -2.435035, -0.737248, 1.570796, 2.395205],accel_mss,speed_ms,0,blend_radius_m)
  movel([0.824257, -1.540869, -2.434309, -0.737211, 1.570796, 2.395053],accel_mss,speed_ms,0,blend_radius_m)
  movel([0.824332, -1.541804, -2.433418, -0.737167, 1.570796, 2.395129],accel_mss,speed_ms,0,blend_radius_m)
  movel([0.824648, -1.542592, -2.432666, -0.737131, 1.570796, 2.395445],accel_mss,speed_ms,0,blend_radius_m)
  movel([0.825204, -1.543233, -2.432054, -0.737103, 1.570796, 2.396000],accel_mss,speed_ms,0,blend_radius_m)
  movel([0.826004, -1.543726, -2.431581, -0.737081, 1.570796, 2.396800],accel_mss,speed_ms,0,blend_radius_m)
  movel([0.826994, -1.544047, -2.431274, -0.737067, 1.570796, 2.397790],accel_mss,speed_ms,0,blend_radius_m)
  movel([0.828132, -1.544165, -2.431161, -0.737062, 1.570796, 2.398928],accel_mss,speed_ms,0,blend_radius_m)
  movel([0.829416, -1.544081, -2.431242, -0.737066, 1.570796, 2.400212],accel_mss,speed_ms,0,blend_radius_m)
  movel([0.830849, -1.543797, -2.431514, -0.737078, 1.570796, 2.401645],accel_mss,speed_ms,0,blend_radius_m)
  movel([0.833262, -1.542886, -2.432384, -0.737118, 1.570796, 2.404058],accel_mss,speed_ms,0,blend_radius_m)
  movel([0.835468, -1.541443, -2.433762, -0.737184, 1.570796, 2.406264],accel_mss,speed_ms,0,blend_radius_m)
  movel([0.836473, -1.540520, -2.434641, -0.737228, 1.570796, 2.407269],accel_mss,speed_ms,0,blend_radius_m)
  movel([0.837382, -1.539466, -2.435643, -0.737280, 1.570796, 2.408179],accel_mss,speed_ms,0,blend_radius_m)
  movel([0.838923, -1.536959, -2.438020, -0.737410, 1.570796, 2.409720],accel_mss,speed_ms,0,blend_radius_m)
  movel([0.840001, -1.533965, -2.440845, -0.737579, 1.570796, 2.410798],accel_mss,speed_ms,0,blend_radius_m)
  movel([0.840521, -1.530536, -2.444064, -0.737789, 1.570796, 2.411318],accel_mss,speed_ms,0,blend_radius_m)
  movel([0.852832, -1.527484, -2.446913, -0.737992, 1.570796, 2.423628],accel_mss,speed_ms,0,blend_radius_m)
  movel([0.851627, -1.542599, -2.432659, -0.737131, 1.570796, 2.422423],accel_mss,speed_ms,0,blend_radius_m)
  movel([0.843729, -1.544510, -2.430831, -0.737048, 1.570796, 2.414525],accel_mss,speed_ms,0,blend_radius_m)
  movel([0.845656, -1.543481, -2.431817, -0.737092, 1.570796, 2.416452],accel_mss,speed_ms,0,blend_radius_m)
  movel([0.847451, -1.542016, -2.433215, -0.737157, 1.570796, 2.418247],accel_mss,speed_ms,0,blend_radius_m)
  movel([0.849020, -1.540188, -2.434957, -0.737244, 1.570796, 2.419817],accel_mss,speed_ms,0,blend_radius_m)
  movel([0.850279, -1.538067, -2.436971, -0.737351, 1.570796, 2.421076],accel_mss,speed_ms,0,blend_radius_m)
  movel([0.851157, -1.535723, -2.439188, -0.737478, 1.570796, 2.421953],accel_mss,speed_ms,0,blend_radius_m)
  movel([0.851585, -1.533237, -2.441530, -0.737622, 1.570796, 2.422381],accel_mss,speed_ms,0,blend_radius_m)
  movel([0.842550, -1.535456, -2.439440, -0.737493, 1.570796, 2.413347],accel_mss,speed_ms,0,blend_radius_m)
  movel([0.842098, -1.538497, -2.436563, -0.737329, 1.570796, 2.412894],accel_mss,speed_ms,0,blend_radius_m)
  movel([0.841163, -1.541524, -2.433684, -0.737180, 1.570796, 2.411959],accel_mss,speed_ms,0,blend_radius_m)
  movel([0.839731, -1.544353, -2.430981, -0.737055, 1.570796, 2.410527],accel_mss,speed_ms,0,blend_radius_m)
  movel([0.838824, -1.545627, -2.429760, -0.737002, 1.570796, 2.409621],accel_mss,speed_ms,0,blend_radius_m)
  movel([0.837787, -1.546808, -2.428625, -0.736956, 1.570796, 2.408583],accel_mss,speed_ms,0,blend_radius_m)
  movel([0.836626, -1.547850, -2.427622, -0.736917, 1.570796, 2.407422],accel_mss,speed_ms,0,blend_radius_m)
  movel([0.835342, -1.548707, -2.426796, -0.736886, 1.570796, 2.406138],accel_mss,speed_ms,0,blend_radius_m)
  movel([0.833934, -1.549383, -2.426144, -0.736863, 1.570796, 2.404731],accel_mss,speed_ms,0,blend_radius_m)
  movel([0.832403, -1.549875, -2.425668, -0.736846, 1.570796, 2.403199],accel_mss,speed_ms,0,blend_radius_m)
  movel([0.830882, -1.550159, -2.425393, -0.736836, 1.570796, 2.401678],accel_mss,speed_ms,0,blend_radius_m)
  movel([0.829503, -1.550212, -2.425343, -0.736835, 1.570796, 2.400299],accel_mss,speed_ms,0,blend_radius_m)
  movel([0.828266, -1.550031, -2.425518, -0.736841, 1.570796, 2.399063],accel_mss,speed_ms,0,blend_radius_m)
  movel([0.827170, -1.549615, -2.425919, -0.736855, 1.570796, 2.397966],accel_mss,speed_ms,0,blend_radius_m)
  movel([0.825405, -1.548264, -2.427223, -0.736902, 1.570796, 2.396202],accel_mss,speed_ms,0,blend_radius_m)
  movel([0.824222, -1.546339, -2.429076, -0.736974, 1.570796, 2.395018],accel_mss,speed_ms,0,blend_radius_m)
  movel([0.823580, -1.544019, -2.431301, -0.737069, 1.570796, 2.394376],accel_mss,speed_ms,0,blend_radius_m)
  movel([0.823445, -1.541489, -2.433718, -0.737182, 1.570796, 2.394241],accel_mss,speed_ms,0,blend_radius_m)
  movel([0.823690, -1.539663, -2.435456, -0.737270, 1.570796, 2.394486],accel_mss,speed_ms,0,blend_radius_m)
  movel([0.824258, -1.537728, -2.437292, -0.737369, 1.570796, 2.395055],accel_mss,speed_ms,0,blend_radius_m)
  movel([0.825132, -1.535855, -2.439063, -0.737470, 1.570796, 2.395929],accel_mss,speed_ms,0,blend_radius_m)
  movel([0.826298, -1.534222, -2.440604, -0.737564, 1.570796, 2.397094],accel_mss,speed_ms,0,blend_radius_m)
  movel([0.827705, -1.532975, -2.441777, -0.737637, 1.570796, 2.398501],accel_mss,speed_ms,0,blend_radius_m)
  movel([0.829309, -1.532262, -2.442446, -0.737681, 1.570796, 2.400105],accel_mss,speed_ms,0,blend_radius_m)
  speed_ms = 0.003
  movel([0.829309, -1.526641, -2.439900, -0.745848, 1.570796, 2.400105],accel_mss,speed_ms,0,blend_radius_m)
  speed_ms = 0.05
  movel([0.829309, -1.504822, -2.429429, -0.778138, 1.570796, 2.400105],accel_mss,speed_ms,0,blend_radius_m)
  #M_RunCode9
  movel([0.860694, -1.432699, -2.490396, -0.789294, 1.570796, 2.431490],accel_mss,speed_ms,0,blend_radius_m)
  #M_RunCode3
  movel([0.860694, -1.456029, -2.501700, -0.754660, 1.570796, 2.431490],accel_mss,speed_ms,0,blend_radius_m)
  speed_ms = 0.003
  movel([0.860694, -1.462060, -2.504453, -0.745876, 1.570796, 2.431490],accel_mss,speed_ms,0,blend_radius_m)
  speed_ms = 0.02
  movel([0.858620, -1.461643, -2.504799, -0.745948, 1.570796, 2.429417],accel_mss,speed_ms,0,blend_radius_m)
  movel([0.856803, -1.460735, -2.505550, -0.746105, 1.570796, 2.427599],accel_mss,speed_ms,0,blend_radius_m)
  movel([0.855243, -1.459441, -2.506618, -0.746330, 1.570796, 2.426040],accel_mss,speed_ms,0,blend_radius_m)
  movel([0.853952, -1.457865, -2.507916, -0.746609, 1.570796, 2.424748],accel_mss,speed_ms,0,blend_radius_m)
  movel([0.852938, -1.456109, -2.509357, -0.746924, 1.570796, 2.423734],accel_mss,speed_ms,0,blend_radius_m)
  movel([0.855159, -1.453688, -2.511335, -0.747365, 1.570796, 2.425956],accel_mss,speed_ms,0,blend_radius_m)
  movel([0.858075, -1.451374, -2.513219, -0.747796, 1.570796, 2.428872],accel_mss,speed_ms,0,blend_radius_m)
  movel([0.861403, -1.449361, -2.514851, -0.748177, 1.570796, 2.432199],accel_mss,speed_ms,0,blend_radius_m)
  movel([0.864838, -1.447853, -2.516069, -0.748467, 1.570796, 2.435635],accel_mss,speed_ms,0,blend_radius_m)
  movel([0.868083, -1.447051, -2.516715, -0.748622, 1.570796, 2.438879],accel_mss,speed_ms,0,blend_radius_m)
  movel([0.869537, -1.446976, -2.516776, -0.748637, 1.570796, 2.440334],accel_mss,speed_ms,0,blend_radius_m)
  movel([0.870830, -1.447150, -2.516636, -0.748603, 1.570796, 2.441627],accel_mss,speed_ms,0,blend_radius_m)
  movel([0.871923, -1.447598, -2.516275, -0.748516, 1.570796, 2.442720],accel_mss,speed_ms,0,blend_radius_m)
  movel([0.872780, -1.448343, -2.515674, -0.748372, 1.570796, 2.443577],accel_mss,speed_ms,0,blend_radius_m)
  movel([0.873364, -1.449404, -2.514816, -0.748169, 1.570796, 2.444160],accel_mss,speed_ms,0,blend_radius_m)
  movel([0.873635, -1.450809, -2.513678, -0.747902, 1.570796, 2.444431],accel_mss,speed_ms,0,blend_radius_m)
  movel([0.873362, -1.453099, -2.511816, -0.747474, 1.570796, 2.444159],accel_mss,speed_ms,0,blend_radius_m)
  movel([0.872321, -1.455315, -2.510006, -0.747067, 1.570796, 2.443117],accel_mss,speed_ms,0,blend_radius_m)
  movel([0.870625, -1.457404, -2.508294, -0.746691, 1.570796, 2.441422],accel_mss,speed_ms,0,blend_radius_m)
  movel([0.868391, -1.459311, -2.506725, -0.746353, 1.570796, 2.439187],accel_mss,speed_ms,0,blend_radius_m)
  movel([0.865580, -1.461003, -2.505328, -0.746058, 1.570796, 2.436377],accel_mss,speed_ms,0,blend_radius_m)
  movel([0.863015, -1.461882, -2.504600, -0.745906, 1.570796, 2.433812],accel_mss,speed_ms,0,blend_radius_m)
  movel([0.860694, -1.462060, -2.504453, -0.745876, 1.570796, 2.431490],accel_mss,speed_ms,0,blend_radius_m)
  speed_ms = 0.003
  movel([0.860694, -1.456029, -2.501700, -0.754660, 1.570796, 2.431490],accel_mss,speed_ms,0,blend_radius_m)
  speed_ms = 0.05
  movel([0.860694, -1.432699, -2.490396, -0.789294, 1.570796, 2.431490],accel_mss,speed_ms,0,blend_radius_m)
  #M_RunCode9
  movel([0.943531, -1.383419, -2.527688, -0.801282, 1.570796, 2.514328],accel_mss,speed_ms,0,blend_radius_m)
  #M_RunCode3
  movel([0.943531, -1.407723, -2.539594, -0.765072, 1.570796, 2.514328],accel_mss,speed_ms,0,blend_radius_m)
  speed_ms = 0.003
  movel([0.943531, -1.414023, -2.542499, -0.755868, 1.570796, 2.514328],accel_mss,speed_ms,0,blend_radius_m)
  speed_ms = 0.02
  movel([0.943228, -1.412692, -2.543503, -0.756194, 1.570796, 2.514024],accel_mss,speed_ms,0,blend_radius_m)
  movel([0.943347, -1.411155, -2.544661, -0.756574, 1.570796, 2.514143],accel_mss,speed_ms,0,blend_radius_m)
  movel([0.943701, -1.409521, -2.545887, -0.756981, 1.570796, 2.514497],accel_mss,speed_ms,0,blend_radius_m)
  movel([0.944289, -1.409603, -2.545825, -0.756961, 1.570796, 2.515085],accel_mss,speed_ms,0,blend_radius_m)
  movel([0.944468, -1.410055, -2.545486, -0.756848, 1.570796, 2.515264],accel_mss,speed_ms,0,blend_radius_m)
  movel([0.944721, -1.410549, -2.545115, -0.756724, 1.570796, 2.515517],accel_mss,speed_ms,0,blend_radius_m)
  movel([0.945526, -1.410758, -2.544958, -0.756672, 1.570796, 2.516322],accel_mss,speed_ms,0,blend_radius_m)
  movel([0.946593, -1.410564, -2.545105, -0.756721, 1.570796, 2.517389],accel_mss,speed_ms,0,blend_radius_m)
  movel([0.947704, -1.410156, -2.545411, -0.756822, 1.570796, 2.518500],accel_mss,speed_ms,0,blend_radius_m)
  movel([0.949249, -1.409535, -2.545876, -0.756978, 1.570796, 2.520045],accel_mss,speed_ms,0,blend_radius_m)
  movel([0.949813, -1.407464, -2.547425, -0.757500, 1.570796, 2.520610],accel_mss,speed_ms,0,blend_radius_m)
  movel([0.949722, -1.405863, -2.548617, -0.757908, 1.570796, 2.520518],accel_mss,speed_ms,0,blend_radius_m)
  movel([0.949358, -1.405315, -2.549025, -0.758049, 1.570796, 2.520154],accel_mss,speed_ms,0,blend_radius_m)
  movel([0.948741, -1.404977, -2.549276, -0.758136, 1.570796, 2.519537],accel_mss,speed_ms,0,blend_radius_m)
  movel([0.947840, -1.404881, -2.549347, -0.758160, 1.570796, 2.518637],accel_mss,speed_ms,0,blend_radius_m)
  movel([0.946628, -1.405061, -2.549214, -0.758114, 1.570796, 2.517424],accel_mss,speed_ms,0,blend_radius_m)
  movel([0.947528, -1.403907, -2.550070, -0.758412, 1.570796, 2.518325],accel_mss,speed_ms,0,blend_radius_m)
  movel([0.948415, -1.402978, -2.550758, -0.758653, 1.570796, 2.519211],accel_mss,speed_ms,0,blend_radius_m)
  movel([0.948839, -1.402709, -2.550957, -0.758723, 1.570796, 2.519635],accel_mss,speed_ms,0,blend_radius_m)
  movel([0.949241, -1.402634, -2.551012, -0.758743, 1.570796, 2.520037],accel_mss,speed_ms,0,blend_radius_m)
  movel([0.949957, -1.403242, -2.550562, -0.758584, 1.570796, 2.520754],accel_mss,speed_ms,0,blend_radius_m)
  movel([0.950638, -1.405149, -2.549149, -0.758092, 1.570796, 2.521435],accel_mss,speed_ms,0,blend_radius_m)
  movel([0.950741, -1.407383, -2.547485, -0.757521, 1.570796, 2.521537],accel_mss,speed_ms,0,blend_radius_m)
  movel([0.950499, -1.408535, -2.546625, -0.757229, 1.570796, 2.521296],accel_mss,speed_ms,0,blend_radius_m)
  movel([0.950018, -1.409665, -2.545779, -0.756945, 1.570796, 2.520814],accel_mss,speed_ms,0,blend_radius_m)
  movel([0.949270, -1.410738, -2.544974, -0.756677, 1.570796, 2.520066],accel_mss,speed_ms,0,blend_radius_m)
  movel([0.948222, -1.411721, -2.544235, -0.756433, 1.570796, 2.519018],accel_mss,speed_ms,0,blend_radius_m)
  movel([0.947736, -1.410561, -2.545107, -0.756721, 1.570796, 2.518532],accel_mss,speed_ms,0,blend_radius_m)
  movel([0.944449, -1.415033, -2.541734, -0.755622, 1.570796, 2.515245],accel_mss,speed_ms,0,blend_radius_m)
  movel([0.943531, -1.414023, -2.542499, -0.755868, 1.570796, 2.514328],accel_mss,speed_ms,0,blend_radius_m)
  speed_ms = 0.003
  movel([0.943531, -1.407723, -2.539594, -0.765072, 1.570796, 2.514328],accel_mss,speed_ms,0,blend_radius_m)
  speed_ms = 0.05
  movel([0.943531, -1.383419, -2.527688, -0.801282, 1.570796, 2.514328],accel_mss,speed_ms,0,blend_radius_m)
  #M_RunCode9
  movel([0.945563, -1.340708, -2.557271, -0.814410, 1.570796, 2.516359],accel_mss,speed_ms,0,blend_radius_m)
  #M_RunCode3
  movel([0.945563, -1.365796, -2.569716, -0.776877, 1.570796, 2.516359],accel_mss,speed_ms,0,blend_radius_m)
  speed_ms = 0.003
  movel([0.945563, -1.372316, -2.572756, -0.767317, 1.570796, 2.516359],accel_mss,speed_ms,0,blend_radius_m)
  speed_ms = 0.02
  movel([0.943258, -1.373056, -2.572241, -0.767092, 1.570796, 2.514055],accel_mss,speed_ms,0,blend_radius_m)
  movel([0.940957, -1.373557, -2.571891, -0.766940, 1.570796, 2.511754],accel_mss,speed_ms,0,blend_radius_m)
  movel([0.938691, -1.373798, -2.571724, -0.766867, 1.570796, 2.509487],accel_mss,speed_ms,0,blend_radius_m)
  movel([0.936487, -1.373762, -2.571749, -0.766878, 1.570796, 2.507284],accel_mss,speed_ms,0,blend_radius_m)
  movel([0.934379, -1.373434, -2.571977, -0.766977, 1.570796, 2.505175],accel_mss,speed_ms,0,blend_radius_m)
  movel([0.933423, -1.373006, -2.572276, -0.767107, 1.570796, 2.504220],accel_mss,speed_ms,0,blend_radius_m)
  movel([0.932562, -1.372371, -2.572717, -0.767300, 1.570796, 2.503358],accel_mss,speed_ms,0,blend_radius_m)
  movel([0.931778, -1.371808, -2.573109, -0.767472, 1.570796, 2.502575],accel_mss,speed_ms,0,blend_radius_m)
  movel([0.931073, -1.371591, -2.573260, -0.767538, 1.570796, 2.501869],accel_mss,speed_ms,0,blend_radius_m)
  movel([0.929539, -1.372029, -2.572956, -0.767405, 1.570796, 2.500335],accel_mss,speed_ms,0,blend_radius_m)
  movel([0.927384, -1.372931, -2.572328, -0.767130, 1.570796, 2.498180],accel_mss,speed_ms,0,blend_radius_m)
  movel([0.925130, -1.373903, -2.571650, -0.766836, 1.570796, 2.495927],accel_mss,speed_ms,0,blend_radius_m)
  movel([0.923297, -1.374547, -2.571201, -0.766641, 1.570796, 2.494093],accel_mss,speed_ms,0,blend_radius_m)
  movel([0.919947, -1.375114, -2.570804, -0.766470, 1.570796, 2.490743],accel_mss,speed_ms,0,blend_radius_m)
  movel([0.917155, -1.375109, -2.570808, -0.766472, 1.570796, 2.487952],accel_mss,speed_ms,0,blend_radius_m)
  movel([0.914870, -1.374586, -2.571174, -0.766630, 1.570796, 2.485667],accel_mss,speed_ms,0,blend_radius_m)
  movel([0.913045, -1.373596, -2.571865, -0.766929, 1.570796, 2.483842],accel_mss,speed_ms,0,blend_radius_m)
  movel([0.911634, -1.372196, -2.572839, -0.767354, 1.570796, 2.482431],accel_mss,speed_ms,0,blend_radius_m)
  movel([0.910594, -1.370436, -2.574061, -0.767892, 1.570796, 2.481391],accel_mss,speed_ms,0,blend_radius_m)
  movel([0.909880, -1.368371, -2.575489, -0.768530, 1.570796, 2.480677],accel_mss,speed_ms,0,blend_radius_m)
  movel([0.909448, -1.366051, -2.577085, -0.769253, 1.570796, 2.480244],accel_mss,speed_ms,0,blend_radius_m)
  movel([0.909251, -1.360875, -2.580620, -0.770894, 1.570796, 2.480047],accel_mss,speed_ms,0,blend_radius_m)
  movel([0.909654, -1.355352, -2.584351, -0.772686, 1.570796, 2.480450],accel_mss,speed_ms,0,blend_radius_m)
  movel([0.910803, -1.345129, -2.591145, -0.776116, 1.570796, 2.481599],accel_mss,speed_ms,0,blend_radius_m)
  movel([0.910870, -1.340748, -2.594012, -0.777629, 1.570796, 2.481667],accel_mss,speed_ms,0,blend_radius_m)
  movel([0.910494, -1.335831, -2.597199, -0.779359, 1.570796, 2.481290],accel_mss,speed_ms,0,blend_radius_m)
  movel([0.909659, -1.330644, -2.600525, -0.781220, 1.570796, 2.480455],accel_mss,speed_ms,0,blend_radius_m)
  movel([0.908357, -1.325460, -2.603814, -0.783115, 1.570796, 2.479153],accel_mss,speed_ms,0,blend_radius_m)
  movel([0.906573, -1.320565, -2.606886, -0.784938, 1.570796, 2.477370],accel_mss,speed_ms,0,blend_radius_m)
  movel([0.904304, -1.316245, -2.609571, -0.786573, 1.570796, 2.475101],accel_mss,speed_ms,0,blend_radius_m)
  movel([0.901546, -1.312796, -2.611697, -0.787897, 1.570796, 2.472342],accel_mss,speed_ms,0,blend_radius_m)
  movel([0.899982, -1.311492, -2.612496, -0.788401, 1.570796, 2.470778],accel_mss,speed_ms,0,blend_radius_m)
  movel([0.898299, -1.310514, -2.613094, -0.788781, 1.570796, 2.469095],accel_mss,speed_ms,0,blend_radius_m)
  movel([0.896342, -1.309794, -2.613534, -0.789061, 1.570796, 2.467138],accel_mss,speed_ms,0,blend_radius_m)
  movel([0.893864, -1.309224, -2.613881, -0.789283, 1.570796, 2.464660],accel_mss,speed_ms,0,blend_radius_m)
  movel([0.890968, -1.308917, -2.614068, -0.789403, 1.570796, 2.461765],accel_mss,speed_ms,0,blend_radius_m)
  movel([0.887766, -1.308975, -2.614033, -0.789381, 1.570796, 2.458562],accel_mss,speed_ms,0,blend_radius_m)
  movel([0.884374, -1.309500, -2.613713, -0.789176, 1.570796, 2.455170],accel_mss,speed_ms,0,blend_radius_m)
  movel([0.880902, -1.310592, -2.613046, -0.788750, 1.570796, 2.451698],accel_mss,speed_ms,0,blend_radius_m)
  movel([0.877469, -1.312349, -2.611971, -0.788069, 1.570796, 2.448266],accel_mss,speed_ms,0,blend_radius_m)
  movel([0.875806, -1.313501, -2.611263, -0.787625, 1.570796, 2.446602],accel_mss,speed_ms,0,blend_radius_m)
  movel([0.874197, -1.314855, -2.610429, -0.787105, 1.570796, 2.444994],accel_mss,speed_ms,0,blend_radius_m)
  movel([0.872040, -1.317227, -2.608963, -0.786200, 1.570796, 2.442836],accel_mss,speed_ms,0,blend_radius_m)
  movel([0.870681, -1.319564, -2.607510, -0.785315, 1.570796, 2.441478],accel_mss,speed_ms,0,blend_radius_m)
  movel([0.870036, -1.321861, -2.606076, -0.784452, 1.570796, 2.440832],accel_mss,speed_ms,0,blend_radius_m)
  movel([0.870021, -1.324109, -2.604665, -0.783615, 1.570796, 2.440817],accel_mss,speed_ms,0,blend_radius_m)
  movel([0.870554, -1.326302, -2.603282, -0.782805, 1.570796, 2.441351],accel_mss,speed_ms,0,blend_radius_m)
  movel([0.871551, -1.328437, -2.601930, -0.782022, 1.570796, 2.442348],accel_mss,speed_ms,0,blend_radius_m)
  movel([0.872933, -1.330508, -2.600612, -0.781269, 1.570796, 2.443729],accel_mss,speed_ms,0,blend_radius_m)
  movel([0.874615, -1.332515, -2.599330, -0.780544, 1.570796, 2.445412],accel_mss,speed_ms,0,blend_radius_m)
  movel([0.878567, -1.336301, -2.596895, -0.779192, 1.570796, 2.449364],accel_mss,speed_ms,0,blend_radius_m)
  movel([0.882785, -1.339748, -2.594662, -0.777978, 1.570796, 2.453582],accel_mss,speed_ms,0,blend_radius_m)
  movel([0.886664, -1.342785, -2.592682, -0.776922, 1.570796, 2.457460],accel_mss,speed_ms,0,blend_radius_m)
  movel([0.889605, -1.345338, -2.591007, -0.776044, 1.570796, 2.460401],accel_mss,speed_ms,0,blend_radius_m)
  movel([0.896251, -1.351902, -2.586659, -0.773827, 1.570796, 2.467048],accel_mss,speed_ms,0,blend_radius_m)
  movel([0.899628, -1.355539, -2.584225, -0.772625, 1.570796, 2.470424],accel_mss,speed_ms,0,blend_radius_m)
  movel([0.901974, -1.358615, -2.582152, -0.771622, 1.570796, 2.472770],accel_mss,speed_ms,0,blend_radius_m)
  movel([0.902641, -1.360004, -2.581211, -0.771174, 1.570796, 2.473437],accel_mss,speed_ms,0,blend_radius_m)
  movel([0.903056, -1.361507, -2.580190, -0.770691, 1.570796, 2.473852],accel_mss,speed_ms,0,blend_radius_m)
  movel([0.903184, -1.364793, -2.577948, -0.769648, 1.570796, 2.473980],accel_mss,speed_ms,0,blend_radius_m)
  movel([0.902480, -1.368343, -2.575508, -0.768538, 1.570796, 2.473277],accel_mss,speed_ms,0,blend_radius_m)
  movel([0.901077, -1.372031, -2.572954, -0.767404, 1.570796, 2.471874],accel_mss,speed_ms,0,blend_radius_m)
  movel([0.899091, -1.375733, -2.570371, -0.766285, 1.570796, 2.469887],accel_mss,speed_ms,0,blend_radius_m)
  movel([0.896639, -1.379334, -2.567840, -0.765215, 1.570796, 2.467435],accel_mss,speed_ms,0,blend_radius_m)
  movel([0.893837, -1.382721, -2.565443, -0.764226, 1.570796, 2.464633],accel_mss,speed_ms,0,blend_radius_m)
  movel([0.890798, -1.385775, -2.563267, -0.763347, 1.570796, 2.461595],accel_mss,speed_ms,0,blend_radius_m)
  movel([0.886743, -1.389087, -2.560891, -0.762410, 1.570796, 2.457539],accel_mss,speed_ms,0,blend_radius_m)
  movel([0.884924, -1.390276, -2.560035, -0.762078, 1.570796, 2.455720],accel_mss,speed_ms,0,blend_radius_m)
  movel([0.883214, -1.391188, -2.559377, -0.761824, 1.570796, 2.454011],accel_mss,speed_ms,0,blend_radius_m)
  movel([0.881598, -1.391853, -2.558896, -0.761640, 1.570796, 2.452395],accel_mss,speed_ms,0,blend_radius_m)
  movel([0.880056, -1.392297, -2.558575, -0.761517, 1.570796, 2.450852],accel_mss,speed_ms,0,blend_radius_m)
  movel([0.877110, -1.392637, -2.558329, -0.761423, 1.570796, 2.447907],accel_mss,speed_ms,0,blend_radius_m)
  movel([0.874230, -1.392421, -2.558485, -0.761483, 1.570796, 2.445026],accel_mss,speed_ms,0,blend_radius_m)
  movel([0.871268, -1.391867, -2.558886, -0.761636, 1.570796, 2.442065],accel_mss,speed_ms,0,blend_radius_m)
  movel([0.864527, -1.390599, -2.559802, -0.761988, 1.570796, 2.435323],accel_mss,speed_ms,0,blend_radius_m)
  movel([0.864160, -1.390572, -2.559822, -0.761995, 1.570796, 2.434956],accel_mss,speed_ms,0,blend_radius_m)
  movel([0.864220, -1.390713, -2.559720, -0.761956, 1.570796, 2.435016],accel_mss,speed_ms,0,blend_radius_m)
  movel([0.865397, -1.391410, -2.559216, -0.761762, 1.570796, 2.436194],accel_mss,speed_ms,0,blend_radius_m)
  movel([0.870411, -1.393867, -2.557436, -0.761086, 1.570796, 2.441207],accel_mss,speed_ms,0,blend_radius_m)
  movel([0.878673, -1.397971, -2.554443, -0.759975, 1.570796, 2.449470],accel_mss,speed_ms,0,blend_radius_m)
  movel([0.872584, -1.398441, -2.554099, -0.759850, 1.570796, 2.443380],accel_mss,speed_ms,0,blend_radius_m)
  movel([0.865922, -1.398637, -2.553955, -0.759797, 1.570796, 2.436718],accel_mss,speed_ms,0,blend_radius_m)
  movel([0.858904, -1.398608, -2.553976, -0.759805, 1.570796, 2.429700],accel_mss,speed_ms,0,blend_radius_m)
  movel([0.851751, -1.398380, -2.554143, -0.759866, 1.570796, 2.422547],accel_mss,speed_ms,0,blend_radius_m)
  movel([0.837922, -1.397458, -2.554818, -0.760113, 1.570796, 2.408718],accel_mss,speed_ms,0,blend_radius_m)
  movel([0.831705, -1.396796, -2.555302, -0.760290, 1.570796, 2.402502],accel_mss,speed_ms,0,blend_radius_m)
  movel([0.826260, -1.396021, -2.555869, -0.760500, 1.570796, 2.397056],accel_mss,speed_ms,0,blend_radius_m)
  movel([0.817080, -1.398428, -2.554108, -0.759853, 1.570796, 2.387876],accel_mss,speed_ms,0,blend_radius_m)
  movel([0.807532, -1.401385, -2.551934, -0.759070, 1.570796, 2.378328],accel_mss,speed_ms,0,blend_radius_m)
  movel([0.787959, -1.408133, -2.546926, -0.757331, 1.570796, 2.358756],accel_mss,speed_ms,0,blend_radius_m)
  movel([0.778218, -1.411521, -2.544385, -0.756483, 1.570796, 2.349015],accel_mss,speed_ms,0,blend_radius_m)
  movel([0.768679, -1.414655, -2.542021, -0.755714, 1.570796, 2.339476],accel_mss,speed_ms,0,blend_radius_m)
  movel([0.759464, -1.417341, -2.539982, -0.755066, 1.570796, 2.330260],accel_mss,speed_ms,0,blend_radius_m)
  movel([0.750683, -1.419383, -2.538425, -0.754581, 1.570796, 2.321479],accel_mss,speed_ms,0,blend_radius_m)
  movel([0.747387, -1.419900, -2.538030, -0.754459, 1.570796, 2.318184],accel_mss,speed_ms,0,blend_radius_m)
  movel([0.744370, -1.420125, -2.537858, -0.754406, 1.570796, 2.315166],accel_mss,speed_ms,0,blend_radius_m)
  movel([0.741646, -1.420066, -2.537903, -0.754420, 1.570796, 2.312443],accel_mss,speed_ms,0,blend_radius_m)
  movel([0.739225, -1.419734, -2.538157, -0.754498, 1.570796, 2.310021],accel_mss,speed_ms,0,blend_radius_m)
  movel([0.737123, -1.419133, -2.538616, -0.754640, 1.570796, 2.307919],accel_mss,speed_ms,0,blend_radius_m)
  movel([0.735352, -1.418270, -2.539275, -0.754844, 1.570796, 2.306148],accel_mss,speed_ms,0,blend_radius_m)
  movel([0.733925, -1.417154, -2.540125, -0.755111, 1.570796, 2.304721],accel_mss,speed_ms,0,blend_radius_m)
  movel([0.732859, -1.415793, -2.541158, -0.755438, 1.570796, 2.303655],accel_mss,speed_ms,0,blend_radius_m)
  movel([0.732170, -1.414190, -2.542372, -0.755827, 1.570796, 2.302966],accel_mss,speed_ms,0,blend_radius_m)
  movel([0.731874, -1.412352, -2.543759, -0.756277, 1.570796, 2.302670],accel_mss,speed_ms,0,blend_radius_m)
  movel([0.731989, -1.410289, -2.545311, -0.756789, 1.570796, 2.302785],accel_mss,speed_ms,0,blend_radius_m)
  movel([0.732529, -1.408005, -2.547021, -0.757363, 1.570796, 2.303325],accel_mss,speed_ms,0,blend_radius_m)
  movel([0.733515, -1.405508, -2.548882, -0.757999, 1.570796, 2.304311],accel_mss,speed_ms,0,blend_radius_m)
  movel([0.734967, -1.402803, -2.550887, -0.758699, 1.570796, 2.305763],accel_mss,speed_ms,0,blend_radius_m)
  movel([0.736902, -1.399898, -2.553029, -0.759462, 1.570796, 2.307698],accel_mss,speed_ms,0,blend_radius_m)
  movel([0.739342, -1.396802, -2.555298, -0.760289, 1.570796, 2.310138],accel_mss,speed_ms,0,blend_radius_m)
  movel([0.740769, -1.398917, -2.553750, -0.759723, 1.570796, 2.311566],accel_mss,speed_ms,0,blend_radius_m)
  movel([0.741550, -1.399879, -2.553043, -0.759467, 1.570796, 2.312347],accel_mss,speed_ms,0,blend_radius_m)
  movel([0.742610, -1.400510, -2.552579, -0.759300, 1.570796, 2.313406],accel_mss,speed_ms,0,blend_radius_m)
  movel([0.743727, -1.400631, -2.552489, -0.759268, 1.570796, 2.314523],accel_mss,speed_ms,0,blend_radius_m)
  movel([0.745263, -1.400459, -2.552616, -0.759314, 1.570796, 2.316059],accel_mss,speed_ms,0,blend_radius_m)
  movel([0.749374, -1.399371, -2.553416, -0.759602, 1.570796, 2.320170],accel_mss,speed_ms,0,blend_radius_m)
  movel([0.754507, -1.397532, -2.554764, -0.760093, 1.570796, 2.325303],accel_mss,speed_ms,0,blend_radius_m)
  movel([0.760223, -1.395214, -2.556456, -0.760718, 1.570796, 2.331019],accel_mss,speed_ms,0,blend_radius_m)
  movel([0.771600, -1.390256, -2.560050, -0.762083, 1.570796, 2.342397],accel_mss,speed_ms,0,blend_radius_m)
  movel([0.779849, -1.386677, -2.562622, -0.763091, 1.570796, 2.350645],accel_mss,speed_ms,0,blend_radius_m)
  movel([0.786938, -1.384123, -2.564445, -0.763821, 1.570796, 2.357734],accel_mss,speed_ms,0,blend_radius_m)
  movel([0.794049, -1.381598, -2.566239, -0.764552, 1.570796, 2.364845],accel_mss,speed_ms,0,blend_radius_m)
  movel([0.783249, -1.378779, -2.568231, -0.765378, 1.570796, 2.354045],accel_mss,speed_ms,0,blend_radius_m)
  movel([0.777784, -1.377033, -2.569460, -0.765896, 1.570796, 2.348580],accel_mss,speed_ms,0,blend_radius_m)
  movel([0.772854, -1.374767, -2.571047, -0.766575, 1.570796, 2.343650],accel_mss,speed_ms,0,blend_radius_m)
  movel([0.770728, -1.373362, -2.572027, -0.766999, 1.570796, 2.341524],accel_mss,speed_ms,0,blend_radius_m)
  movel([0.768902, -1.371738, -2.573158, -0.767494, 1.570796, 2.339698],accel_mss,speed_ms,0,blend_radius_m)
  movel([0.767434, -1.369859, -2.574461, -0.768070, 1.570796, 2.338230],accel_mss,speed_ms,0,blend_radius_m)
  movel([0.766379, -1.367694, -2.575955, -0.768740, 1.570796, 2.337175],accel_mss,speed_ms,0,blend_radius_m)
  movel([0.765796, -1.365211, -2.577661, -0.769517, 1.570796, 2.336592],accel_mss,speed_ms,0,blend_radius_m)
  movel([0.765745, -1.362374, -2.579600, -0.770415, 1.570796, 2.336542],accel_mss,speed_ms,0,blend_radius_m)
  movel([0.766289, -1.359146, -2.581793, -0.771451, 1.570796, 2.337086],accel_mss,speed_ms,0,blend_radius_m)
  movel([0.767492, -1.355492, -2.584257, -0.772640, 1.570796, 2.338288],accel_mss,speed_ms,0,blend_radius_m)
  movel([0.769653, -1.351141, -2.587167, -0.774081, 1.570796, 2.340450],accel_mss,speed_ms,0,blend_radius_m)
  movel([0.772614, -1.346772, -2.590062, -0.775555, 1.570796, 2.343411],accel_mss,speed_ms,0,blend_radius_m)
  movel([0.776249, -1.342511, -2.592861, -0.777017, 1.570796, 2.347045],accel_mss,speed_ms,0,blend_radius_m)
  movel([0.780428, -1.338491, -2.595479, -0.778419, 1.570796, 2.351224],accel_mss,speed_ms,0,blend_radius_m)
  movel([0.785012, -1.334851, -2.597830, -0.779708, 1.570796, 2.355808],accel_mss,speed_ms,0,blend_radius_m)
  movel([0.789857, -1.331729, -2.599832, -0.780827, 1.570796, 2.360653],accel_mss,speed_ms,0,blend_radius_m)
  movel([0.794818, -1.329265, -2.601404, -0.781720, 1.570796, 2.365614],accel_mss,speed_ms,0,blend_radius_m)
  movel([0.799737, -1.327602, -2.602460, -0.782328, 1.570796, 2.370534],accel_mss,speed_ms,0,blend_radius_m)
  movel([0.802223, -1.327350, -2.602619, -0.782420, 1.570796, 2.373019],accel_mss,speed_ms,0,blend_radius_m)
  movel([0.804703, -1.327682, -2.602409, -0.782298, 1.570796, 2.375499],accel_mss,speed_ms,0,blend_radius_m)
  movel([0.806357, -1.328539, -2.601865, -0.781985, 1.570796, 2.377153],accel_mss,speed_ms,0,blend_radius_m)
  movel([0.806622, -1.329147, -2.601479, -0.781763, 1.570796, 2.377418],accel_mss,speed_ms,0,blend_radius_m)
  movel([0.806375, -1.329863, -2.601023, -0.781503, 1.570796, 2.377171],accel_mss,speed_ms,0,blend_radius_m)
  movel([0.804438, -1.329565, -2.601213, -0.781611, 1.570796, 2.375234],accel_mss,speed_ms,0,blend_radius_m)
  movel([0.802662, -1.329558, -2.601217, -0.781614, 1.570796, 2.373458],accel_mss,speed_ms,0,blend_radius_m)
  movel([0.801050, -1.329817, -2.601052, -0.781519, 1.570796, 2.371846],accel_mss,speed_ms,0,blend_radius_m)
  movel([0.799606, -1.330312, -2.600737, -0.781340, 1.570796, 2.370402],accel_mss,speed_ms,0,blend_radius_m)
  movel([0.798332, -1.331017, -2.600288, -0.781085, 1.570796, 2.369129],accel_mss,speed_ms,0,blend_radius_m)
  movel([0.797239, -1.331898, -2.599725, -0.780766, 1.570796, 2.368035],accel_mss,speed_ms,0,blend_radius_m)
  movel([0.796324, -1.332932, -2.599063, -0.780395, 1.570796, 2.367121],accel_mss,speed_ms,0,blend_radius_m)
  movel([0.795591, -1.334089, -2.598320, -0.779980, 1.570796, 2.366387],accel_mss,speed_ms,0,blend_radius_m)
  movel([0.794681, -1.336663, -2.596662, -0.779064, 1.570796, 2.365478],accel_mss,speed_ms,0,blend_radius_m)
  movel([0.794525, -1.339402, -2.594888, -0.778099, 1.570796, 2.365322],accel_mss,speed_ms,0,blend_radius_m)
  movel([0.795140, -1.342094, -2.593134, -0.777161, 1.570796, 2.365937],accel_mss,speed_ms,0,blend_radius_m)
  movel([0.796533, -1.344536, -2.591534, -0.776319, 1.570796, 2.367330],accel_mss,speed_ms,0,blend_radius_m)
  movel([0.797751, -1.345705, -2.590766, -0.775919, 1.570796, 2.368548],accel_mss,speed_ms,0,blend_radius_m)
  movel([0.799475, -1.346850, -2.590011, -0.775528, 1.570796, 2.370271],accel_mss,speed_ms,0,blend_radius_m)
  movel([0.804179, -1.349059, -2.588550, -0.774780, 1.570796, 2.374975],accel_mss,speed_ms,0,blend_radius_m)
  movel([0.810111, -1.351157, -2.587156, -0.774076, 1.570796, 2.380907],accel_mss,speed_ms,0,blend_radius_m)
  movel([0.816751, -1.353123, -2.585844, -0.773422, 1.570796, 2.387547],accel_mss,speed_ms,0,blend_radius_m)
  movel([0.830115, -1.356522, -2.583564, -0.772303, 1.570796, 2.400912],accel_mss,speed_ms,0,blend_radius_m)
  movel([0.840314, -1.358817, -2.582015, -0.771557, 1.570796, 2.411110],accel_mss,speed_ms,0,blend_radius_m)
  movel([0.845440, -1.359957, -2.581243, -0.771189, 1.570796, 2.416236],accel_mss,speed_ms,0,blend_radius_m)
  movel([0.848261, -1.360460, -2.580902, -0.771027, 1.570796, 2.419057],accel_mss,speed_ms,0,blend_radius_m)
  movel([0.850527, -1.360613, -2.580798, -0.770978, 1.570796, 2.421323],accel_mss,speed_ms,0,blend_radius_m)
  movel([0.851222, -1.360500, -2.580875, -0.771014, 1.570796, 2.422018],accel_mss,speed_ms,0,blend_radius_m)
  movel([0.851602, -1.360246, -2.581047, -0.771096, 1.570796, 2.422398],accel_mss,speed_ms,0,blend_radius_m)
  movel([0.851751, -1.359254, -2.581720, -0.771416, 1.570796, 2.422547],accel_mss,speed_ms,0,blend_radius_m)
  movel([0.851172, -1.356700, -2.583444, -0.772245, 1.570796, 2.421968],accel_mss,speed_ms,0,blend_radius_m)
  movel([0.850009, -1.354369, -2.585010, -0.773010, 1.570796, 2.420805],accel_mss,speed_ms,0,blend_radius_m)
  movel([0.847204, -1.349555, -2.588221, -0.774613, 1.570796, 2.418000],accel_mss,speed_ms,0,blend_radius_m)
  movel([0.846203, -1.346648, -2.590144, -0.775597, 1.570796, 2.416999],accel_mss,speed_ms,0,blend_radius_m)
  movel([0.845909, -1.343110, -2.592469, -0.776810, 1.570796, 2.416705],accel_mss,speed_ms,0,blend_radius_m)
  movel([0.846133, -1.341034, -2.593825, -0.777530, 1.570796, 2.416929],accel_mss,speed_ms,0,blend_radius_m)
  movel([0.846657, -1.338714, -2.595334, -0.778341, 1.570796, 2.417454],accel_mss,speed_ms,0,blend_radius_m)
  movel([0.847529, -1.336119, -2.597013, -0.779257, 1.570796, 2.418326],accel_mss,speed_ms,0,blend_radius_m)
  movel([0.848795, -1.333217, -2.598880, -0.780292, 1.570796, 2.419591],accel_mss,speed_ms,0,blend_radius_m)
  movel([0.850964, -1.329406, -2.601314, -0.781669, 1.570796, 2.421760],accel_mss,speed_ms,0,blend_radius_m)
  movel([0.853600, -1.325900, -2.603536, -0.782953, 1.570796, 2.424397],accel_mss,speed_ms,0,blend_radius_m)
  movel([0.856646, -1.322679, -2.605563, -0.784147, 1.570796, 2.427443],accel_mss,speed_ms,0,blend_radius_m)
  movel([0.860034, -1.319733, -2.607405, -0.785251, 1.570796, 2.430830],accel_mss,speed_ms,0,blend_radius_m)
  movel([0.863699, -1.317039, -2.609079, -0.786271, 1.570796, 2.434495],accel_mss,speed_ms,0,blend_radius_m)
  movel([0.867570, -1.314582, -2.610598, -0.787209, 1.570796, 2.438367],accel_mss,speed_ms,0,blend_radius_m)
  movel([0.871586, -1.312340, -2.611976, -0.788073, 1.570796, 2.442383],accel_mss,speed_ms,0,blend_radius_m)
  movel([0.875674, -1.310295, -2.613228, -0.788866, 1.570796, 2.446470],accel_mss,speed_ms,0,blend_radius_m)
  movel([0.883349, -1.307075, -2.615188, -0.790126, 1.570796, 2.454145],accel_mss,speed_ms,0,blend_radius_m)
  movel([0.889958, -1.305028, -2.616427, -0.790934, 1.570796, 2.460755],accel_mss,speed_ms,0,blend_radius_m)
  movel([0.895338, -1.303917, -2.617097, -0.791375, 1.570796, 2.466135],accel_mss,speed_ms,0,blend_radius_m)
  movel([0.899336, -1.303497, -2.617350, -0.791542, 1.570796, 2.470133],accel_mss,speed_ms,0,blend_radius_m)
  movel([0.904889, -1.303658, -2.617253, -0.791478, 1.570796, 2.475686],accel_mss,speed_ms,0,blend_radius_m)
  movel([0.909830, -1.304667, -2.616645, -0.791077, 1.570796, 2.480626],accel_mss,speed_ms,0,blend_radius_m)
  movel([0.914127, -1.306464, -2.615559, -0.790367, 1.570796, 2.484923],accel_mss,speed_ms,0,blend_radius_m)
  movel([0.917751, -1.308972, -2.614035, -0.789382, 1.570796, 2.488547],accel_mss,speed_ms,0,blend_radius_m)
  movel([0.920676, -1.312123, -2.612109, -0.788156, 1.570796, 2.491473],accel_mss,speed_ms,0,blend_radius_m)
  movel([0.922887, -1.315842, -2.609820, -0.786727, 1.570796, 2.493683],accel_mss,speed_ms,0,blend_radius_m)
  movel([0.924365, -1.320052, -2.607206, -0.785131, 1.570796, 2.495162],accel_mss,speed_ms,0,blend_radius_m)
  movel([0.925096, -1.324684, -2.604303, -0.783402, 1.570796, 2.495892],accel_mss,speed_ms,0,blend_radius_m)
  movel([0.925102, -1.329152, -2.601476, -0.781762, 1.570796, 2.495899],accel_mss,speed_ms,0,blend_radius_m)
  movel([0.924715, -1.333726, -2.598553, -0.780110, 1.570796, 2.495512],accel_mss,speed_ms,0,blend_radius_m)
  movel([0.924273, -1.338230, -2.595648, -0.778511, 1.570796, 2.495069],accel_mss,speed_ms,0,blend_radius_m)
  movel([0.924113, -1.342493, -2.592873, -0.777023, 1.570796, 2.494909],accel_mss,speed_ms,0,blend_radius_m)
  movel([0.924559, -1.346357, -2.590336, -0.775696, 1.570796, 2.495355],accel_mss,speed_ms,0,blend_radius_m)
  movel([0.925111, -1.348086, -2.589194, -0.775109, 1.570796, 2.495908],accel_mss,speed_ms,0,blend_radius_m)
  movel([0.925934, -1.349657, -2.588153, -0.774579, 1.570796, 2.496730],accel_mss,speed_ms,0,blend_radius_m)
  movel([0.927068, -1.351051, -2.587227, -0.774111, 1.570796, 2.497864],accel_mss,speed_ms,0,blend_radius_m)
  movel([0.928552, -1.352249, -2.586428, -0.773712, 1.570796, 2.499348],accel_mss,speed_ms,0,blend_radius_m)
  movel([0.930429, -1.353235, -2.585770, -0.773385, 1.570796, 2.501225],accel_mss,speed_ms,0,blend_radius_m)
  movel([0.932737, -1.353987, -2.585266, -0.773136, 1.570796, 2.503533],accel_mss,speed_ms,0,blend_radius_m)
  movel([0.935000, -1.354278, -2.585072, -0.773040, 1.570796, 2.505796],accel_mss,speed_ms,0,blend_radius_m)
  movel([0.937183, -1.354056, -2.585220, -0.773113, 1.570796, 2.507979],accel_mss,speed_ms,0,blend_radius_m)
  movel([0.939253, -1.353395, -2.585663, -0.773332, 1.570796, 2.510049],accel_mss,speed_ms,0,blend_radius_m)
  movel([0.941181, -1.352368, -2.586349, -0.773672, 1.570796, 2.511977],accel_mss,speed_ms,0,blend_radius_m)
  movel([0.942932, -1.351044, -2.587231, -0.774114, 1.570796, 2.513729],accel_mss,speed_ms,0,blend_radius_m)
  movel([0.944471, -1.349497, -2.588259, -0.774633, 1.570796, 2.515267],accel_mss,speed_ms,0,blend_radius_m)
  movel([0.945765, -1.347801, -2.589382, -0.775205, 1.570796, 2.516561],accel_mss,speed_ms,0,blend_radius_m)
  movel([0.946776, -1.346030, -2.590552, -0.775808, 1.570796, 2.517573],accel_mss,speed_ms,0,blend_radius_m)
  movel([0.947469, -1.344259, -2.591716, -0.776414, 1.570796, 2.518265],accel_mss,speed_ms,0,blend_radius_m)
  movel([0.947803, -1.342564, -2.592826, -0.776998, 1.570796, 2.518599],accel_mss,speed_ms,0,blend_radius_m)
  movel([0.947740, -1.341025, -2.593832, -0.777533, 1.570796, 2.518537],accel_mss,speed_ms,0,blend_radius_m)
  movel([0.947242, -1.339719, -2.594682, -0.777989, 1.570796, 2.518039],accel_mss,speed_ms,0,blend_radius_m)
  movel([0.946274, -1.338721, -2.595329, -0.778338, 1.570796, 2.517071],accel_mss,speed_ms,0,blend_radius_m)
  movel([0.944796, -1.338119, -2.595720, -0.778550, 1.570796, 2.515592],accel_mss,speed_ms,0,blend_radius_m)
  movel([0.942768, -1.337990, -2.595804, -0.778596, 1.570796, 2.513565],accel_mss,speed_ms,0,blend_radius_m)
  movel([0.940162, -1.338409, -2.595532, -0.778448, 1.570796, 2.510958],accel_mss,speed_ms,0,blend_radius_m)
  movel([0.941066, -1.339371, -2.594908, -0.778110, 1.570796, 2.511863],accel_mss,speed_ms,0,blend_radius_m)
  movel([0.941537, -1.340439, -2.594213, -0.777737, 1.570796, 2.512334],accel_mss,speed_ms,0,blend_radius_m)
  movel([0.941591, -1.341564, -2.593480, -0.777345, 1.570796, 2.512387],accel_mss,speed_ms,0,blend_radius_m)
  movel([0.941243, -1.342699, -2.592738, -0.776952, 1.570796, 2.512039],accel_mss,speed_ms,0,blend_radius_m)
  movel([0.940505, -1.343800, -2.592017, -0.776572, 1.570796, 2.511302],accel_mss,speed_ms,0,blend_radius_m)
  movel([0.939394, -1.344820, -2.591348, -0.776222, 1.570796, 2.510190],accel_mss,speed_ms,0,blend_radius_m)
  movel([0.937924, -1.345711, -2.590761, -0.775916, 1.570796, 2.508721],accel_mss,speed_ms,0,blend_radius_m)
  movel([0.936108, -1.346430, -2.590288, -0.775671, 1.570796, 2.506904],accel_mss,speed_ms,0,blend_radius_m)
  movel([0.933072, -1.347044, -2.589883, -0.775462, 1.570796, 2.503869],accel_mss,speed_ms,0,blend_radius_m)
  movel([0.930629, -1.346865, -2.590001, -0.775523, 1.570796, 2.501425],accel_mss,speed_ms,0,blend_radius_m)
  movel([0.928748, -1.345988, -2.590579, -0.775822, 1.570796, 2.499544],accel_mss,speed_ms,0,blend_radius_m)
  movel([0.927414, -1.344511, -2.591550, -0.776327, 1.570796, 2.498210],accel_mss,speed_ms,0,blend_radius_m)
  movel([0.926608, -1.342525, -2.592852, -0.777012, 1.570796, 2.497405],accel_mss,speed_ms,0,blend_radius_m)
  movel([0.926317, -1.340123, -2.594419, -0.777847, 1.570796, 2.497113],accel_mss,speed_ms,0,blend_radius_m)
  movel([0.926527, -1.337402, -2.596184, -0.778803, 1.570796, 2.497324],accel_mss,speed_ms,0,blend_radius_m)
  movel([0.927221, -1.334456, -2.598084, -0.779849, 1.570796, 2.498018],accel_mss,speed_ms,0,blend_radius_m)
  movel([0.928394, -1.331380, -2.600056, -0.780953, 1.570796, 2.499190],accel_mss,speed_ms,0,blend_radius_m)
  movel([0.930022, -1.328277, -2.602031, -0.782081, 1.570796, 2.500818],accel_mss,speed_ms,0,blend_radius_m)
  movel([0.932099, -1.325245, -2.603949, -0.783194, 1.570796, 2.502895],accel_mss,speed_ms,0,blend_radius_m)
  movel([0.934601, -1.322396, -2.605741, -0.784253, 1.570796, 2.505397],accel_mss,speed_ms,0,blend_radius_m)
  movel([0.937516, -1.319830, -2.607344, -0.785214, 1.570796, 2.508312],accel_mss,speed_ms,0,blend_radius_m)
  movel([0.940819, -1.317661, -2.608693, -0.786034, 1.570796, 2.511615],accel_mss,speed_ms,0,blend_radius_m)
  movel([0.944488, -1.316003, -2.609720, -0.786666, 1.570796, 2.515284],accel_mss,speed_ms,0,blend_radius_m)
  movel([0.948495, -1.314966, -2.610361, -0.787062, 1.570796, 2.519291],accel_mss,speed_ms,0,blend_radius_m)
  movel([0.951289, -1.314634, -2.610566, -0.787189, 1.570796, 2.522085],accel_mss,speed_ms,0,blend_radius_m)
  movel([0.953948, -1.314579, -2.610599, -0.787211, 1.570796, 2.524744],accel_mss,speed_ms,0,blend_radius_m)
  movel([0.956456, -1.314785, -2.610473, -0.787132, 1.570796, 2.527252],accel_mss,speed_ms,0,blend_radius_m)
  movel([0.958792, -1.315252, -2.610184, -0.786953, 1.570796, 2.529588],accel_mss,speed_ms,0,blend_radius_m)
  movel([0.960938, -1.315966, -2.609743, -0.786680, 1.570796, 2.531735],accel_mss,speed_ms,0,blend_radius_m)
  movel([0.962879, -1.316922, -2.609152, -0.786316, 1.570796, 2.533675],accel_mss,speed_ms,0,blend_radius_m)
  movel([0.964594, -1.318109, -2.608415, -0.785865, 1.570796, 2.535391],accel_mss,speed_ms,0,blend_radius_m)
  movel([0.966072, -1.319515, -2.607541, -0.785333, 1.570796, 2.536868],accel_mss,speed_ms,0,blend_radius_m)
  movel([0.967291, -1.321132, -2.606532, -0.784725, 1.570796, 2.538088],accel_mss,speed_ms,0,blend_radius_m)
  movel([0.968242, -1.322947, -2.605395, -0.784047, 1.570796, 2.539038],accel_mss,speed_ms,0,blend_radius_m)
  movel([0.968904, -1.324954, -2.604133, -0.783302, 1.570796, 2.539700],accel_mss,speed_ms,0,blend_radius_m)
  movel([0.969266, -1.327140, -2.602752, -0.782497, 1.570796, 2.540062],accel_mss,speed_ms,0,blend_radius_m)
  movel([0.969312, -1.329494, -2.601258, -0.781637, 1.570796, 2.540108],accel_mss,speed_ms,0,blend_radius_m)
  movel([0.969033, -1.332004, -2.599656, -0.780728, 1.570796, 2.539829],accel_mss,speed_ms,0,blend_radius_m)
  movel([0.968409, -1.334664, -2.597951, -0.779775, 1.570796, 2.539205],accel_mss,speed_ms,0,blend_radius_m)
  movel([0.967431, -1.337461, -2.596146, -0.778782, 1.570796, 2.538227],accel_mss,speed_ms,0,blend_radius_m)
  movel([0.965854, -1.340244, -2.594340, -0.777805, 1.570796, 2.536651],accel_mss,speed_ms,0,blend_radius_m)
  movel([0.963680, -1.343183, -2.592421, -0.776785, 1.570796, 2.534476],accel_mss,speed_ms,0,blend_radius_m)
  movel([0.961694, -1.345676, -2.590784, -0.775928, 1.570796, 2.532491],accel_mss,speed_ms,0,blend_radius_m)
  movel([0.960671, -1.347129, -2.589827, -0.775433, 1.570796, 2.531467],accel_mss,speed_ms,0,blend_radius_m)
  movel([0.960755, -1.348217, -2.589107, -0.775064, 1.570796, 2.531552],accel_mss,speed_ms,0,blend_radius_m)
  movel([0.961316, -1.349785, -2.588068, -0.774536, 1.570796, 2.532113],accel_mss,speed_ms,0,blend_radius_m)
  movel([0.961937, -1.351511, -2.586920, -0.773958, 1.570796, 2.532733],accel_mss,speed_ms,0,blend_radius_m)
  movel([0.962208, -1.353066, -2.585882, -0.773441, 1.570796, 2.533004],accel_mss,speed_ms,0,blend_radius_m)
  movel([0.961954, -1.355348, -2.584353, -0.772688, 1.570796, 2.532750],accel_mss,speed_ms,0,blend_radius_m)
  movel([0.961348, -1.357576, -2.582854, -0.771960, 1.570796, 2.532144],accel_mss,speed_ms,0,blend_radius_m)
  movel([0.960421, -1.359731, -2.581396, -0.771262, 1.570796, 2.531217],accel_mss,speed_ms,0,blend_radius_m)
  movel([0.959210, -1.361796, -2.579994, -0.770599, 1.570796, 2.530006],accel_mss,speed_ms,0,blend_radius_m)
  movel([0.957748, -1.363756, -2.578657, -0.769976, 1.570796, 2.528544],accel_mss,speed_ms,0,blend_radius_m)
  movel([0.956070, -1.365589, -2.577402, -0.769398, 1.570796, 2.526866],accel_mss,speed_ms,0,blend_radius_m)
  movel([0.954209, -1.367283, -2.576238, -0.768868, 1.570796, 2.525005],accel_mss,speed_ms,0,blend_radius_m)
  movel([0.952196, -1.368818, -2.575180, -0.768391, 1.570796, 2.522993],accel_mss,speed_ms,0,blend_radius_m)
  movel([0.950062, -1.370181, -2.574237, -0.767971, 1.570796, 2.520859],accel_mss,speed_ms,0,blend_radius_m)
  movel([0.947842, -1.371352, -2.573426, -0.767611, 1.570796, 2.518638],accel_mss,speed_ms,0,blend_radius_m)
  movel([0.945563, -1.372316, -2.572756, -0.767317, 1.570796, 2.516359],accel_mss,speed_ms,0,blend_radius_m)
  speed_ms = 0.003
  movel([0.945563, -1.365796, -2.569716, -0.776877, 1.570796, 2.516359],accel_mss,speed_ms,0,blend_radius_m)
  speed_ms = 0.05
  movel([0.945563, -1.340708, -2.557271, -0.814410, 1.570796, 2.516359],accel_mss,speed_ms,0,blend_radius_m)
  #M_RunCode9
  movel([0.956193, -1.345931, -2.553786, -0.812673, 1.570796, 2.526990],accel_mss,speed_ms,0,blend_radius_m)
  #M_RunCode3
  movel([0.956193, -1.370927, -2.566164, -0.775298, 1.570796, 2.526990],accel_mss,speed_ms,0,blend_radius_m)
  speed_ms = 0.003
  movel([0.956193, -1.377420, -2.569187, -0.765781, 1.570796, 2.526990],accel_mss,speed_ms,0,blend_radius_m)
  speed_ms = 0.02
  movel([0.957569, -1.375878, -2.570269, -0.766241, 1.570796, 2.528365],accel_mss,speed_ms,0,blend_radius_m)
  movel([0.960713, -1.372951, -2.572314, -0.767124, 1.570796, 2.531509],accel_mss,speed_ms,0,blend_radius_m)
  movel([0.963663, -1.370019, -2.574350, -0.768021, 1.570796, 2.534459],accel_mss,speed_ms,0,blend_radius_m)
  movel([0.964794, -1.368470, -2.575420, -0.768499, 1.570796, 2.535591],accel_mss,speed_ms,0,blend_radius_m)
  movel([0.965552, -1.366818, -2.576558, -0.769013, 1.570796, 2.536349],accel_mss,speed_ms,0,blend_radius_m)
  movel([0.965393, -1.367989, -2.575752, -0.768648, 1.570796, 2.536190],accel_mss,speed_ms,0,blend_radius_m)
  movel([0.964673, -1.370171, -2.574244, -0.767974, 1.570796, 2.535469],accel_mss,speed_ms,0,blend_radius_m)
  movel([0.963528, -1.372163, -2.572862, -0.767364, 1.570796, 2.534324],accel_mss,speed_ms,0,blend_radius_m)
  movel([0.962090, -1.374027, -2.571564, -0.766798, 1.570796, 2.532886],accel_mss,speed_ms,0,blend_radius_m)
  movel([0.960489, -1.375823, -2.570308, -0.766258, 1.570796, 2.531285],accel_mss,speed_ms,0,blend_radius_m)
  movel([0.957315, -1.379451, -2.567758, -0.765180, 1.570796, 2.528112],accel_mss,speed_ms,0,blend_radius_m)
  movel([0.955999, -1.381401, -2.566379, -0.764609, 1.570796, 2.526796],accel_mss,speed_ms,0,blend_radius_m)
  movel([0.955038, -1.383515, -2.564878, -0.763996, 1.570796, 2.525834],accel_mss,speed_ms,0,blend_radius_m)
  movel([0.954416, -1.385883, -2.563190, -0.763317, 1.570796, 2.525212],accel_mss,speed_ms,0,blend_radius_m)
  movel([0.954206, -1.387128, -2.562298, -0.762963, 1.570796, 2.525002],accel_mss,speed_ms,0,blend_radius_m)
  movel([0.954262, -1.387805, -2.561813, -0.762771, 1.570796, 2.525058],accel_mss,speed_ms,0,blend_radius_m)
  movel([0.955348, -1.387862, -2.561772, -0.762755, 1.570796, 2.526144],accel_mss,speed_ms,0,blend_radius_m)
  movel([0.956212, -1.387957, -2.561704, -0.762728, 1.570796, 2.527009],accel_mss,speed_ms,0,blend_radius_m)
  movel([0.956988, -1.388243, -2.561499, -0.762648, 1.570796, 2.527785],accel_mss,speed_ms,0,blend_radius_m)
  movel([0.958190, -1.389200, -2.560810, -0.762378, 1.570796, 2.528986],accel_mss,speed_ms,0,blend_radius_m)
  movel([0.958837, -1.390170, -2.560112, -0.762107, 1.570796, 2.529634],accel_mss,speed_ms,0,blend_radius_m)
  movel([0.959044, -1.391165, -2.559394, -0.761830, 1.570796, 2.529841],accel_mss,speed_ms,0,blend_radius_m)
  movel([0.958920, -1.392210, -2.558638, -0.761541, 1.570796, 2.529716],accel_mss,speed_ms,0,blend_radius_m)
  movel([0.958114, -1.394531, -2.556953, -0.760904, 1.570796, 2.528910],accel_mss,speed_ms,0,blend_radius_m)
  movel([0.957293, -1.397305, -2.554931, -0.760154, 1.570796, 2.528089],accel_mss,speed_ms,0,blend_radius_m)
  movel([0.956833, -1.400924, -2.552274, -0.759191, 1.570796, 2.527629],accel_mss,speed_ms,0,blend_radius_m)
  movel([0.956526, -1.404475, -2.549649, -0.758265, 1.570796, 2.527322],accel_mss,speed_ms,0,blend_radius_m)
  movel([0.956042, -1.408049, -2.546988, -0.757352, 1.570796, 2.526838],accel_mss,speed_ms,0,blend_radius_m)
  movel([0.955067, -1.411725, -2.544232, -0.756432, 1.570796, 2.525864],accel_mss,speed_ms,0,blend_radius_m)
  movel([0.954226, -1.413740, -2.542712, -0.755937, 1.570796, 2.525022],accel_mss,speed_ms,0,blend_radius_m)
  movel([0.953174, -1.415734, -2.541203, -0.755452, 1.570796, 2.523970],accel_mss,speed_ms,0,blend_radius_m)
  movel([0.950663, -1.419654, -2.538219, -0.754517, 1.570796, 2.521459],accel_mss,speed_ms,0,blend_radius_m)
  movel([0.947979, -1.423474, -2.535288, -0.753627, 1.570796, 2.518775],accel_mss,speed_ms,0,blend_radius_m)
  movel([0.945568, -1.427175, -2.532428, -0.752786, 1.570796, 2.516364],accel_mss,speed_ms,0,blend_radius_m)
  movel([0.942301, -1.433384, -2.527584, -0.751421, 1.570796, 2.513098],accel_mss,speed_ms,0,blend_radius_m)
  movel([0.940979, -1.436039, -2.525494, -0.750855, 1.570796, 2.511776],accel_mss,speed_ms,0,blend_radius_m)
  movel([0.939580, -1.438519, -2.523533, -0.750336, 1.570796, 2.510376],accel_mss,speed_ms,0,blend_radius_m)
  movel([0.937900, -1.440918, -2.521628, -0.749843, 1.570796, 2.508696],accel_mss,speed_ms,0,blend_radius_m)
  movel([0.935730, -1.443326, -2.519706, -0.749357, 1.570796, 2.506526],accel_mss,speed_ms,0,blend_radius_m)
  movel([0.932865, -1.445836, -2.517693, -0.748860, 1.570796, 2.503662],accel_mss,speed_ms,0,blend_radius_m)
  movel([0.929109, -1.448540, -2.515515, -0.748334, 1.570796, 2.499905],accel_mss,speed_ms,0,blend_radius_m)
  movel([0.925915, -1.450502, -2.513927, -0.747960, 1.570796, 2.496712],accel_mss,speed_ms,0,blend_radius_m)
  movel([0.922885, -1.452056, -2.512665, -0.747668, 1.570796, 2.493681],accel_mss,speed_ms,0,blend_radius_m)
  movel([0.920010, -1.453227, -2.511712, -0.747450, 1.570796, 2.490807],accel_mss,speed_ms,0,blend_radius_m)
  movel([0.917281, -1.454037, -2.511051, -0.747301, 1.570796, 2.488077],accel_mss,speed_ms,0,blend_radius_m)
  movel([0.914694, -1.454513, -2.510662, -0.747214, 1.570796, 2.485490],accel_mss,speed_ms,0,blend_radius_m)
  movel([0.912242, -1.454674, -2.510531, -0.747184, 1.570796, 2.483038],accel_mss,speed_ms,0,blend_radius_m)
  movel([0.909922, -1.454543, -2.510638, -0.747208, 1.570796, 2.480718],accel_mss,speed_ms,0,blend_radius_m)
  movel([0.907727, -1.454140, -2.510967, -0.747282, 1.570796, 2.478523],accel_mss,speed_ms,0,blend_radius_m)
  movel([0.905656, -1.453488, -2.511499, -0.747402, 1.570796, 2.476453],accel_mss,speed_ms,0,blend_radius_m)
  movel([0.903702, -1.452607, -2.512217, -0.747565, 1.570796, 2.474499],accel_mss,speed_ms,0,blend_radius_m)
  movel([0.900139, -1.450236, -2.514142, -0.748011, 1.570796, 2.470935],accel_mss,speed_ms,0,blend_radius_m)
  movel([0.897015, -1.447193, -2.516601, -0.748595, 1.570796, 2.467812],accel_mss,speed_ms,0,blend_radius_m)
  movel([0.894312, -1.443643, -2.519453, -0.749294, 1.570796, 2.465108],accel_mss,speed_ms,0,blend_radius_m)
  movel([0.892214, -1.439938, -2.522408, -0.750044, 1.570796, 2.463010],accel_mss,speed_ms,0,blend_radius_m)
  movel([0.889634, -1.435087, -2.526245, -0.751057, 1.570796, 2.460430],accel_mss,speed_ms,0,blend_radius_m)
  movel([0.886430, -1.429922, -2.530292, -0.752175, 1.570796, 2.457227],accel_mss,speed_ms,0,blend_radius_m)
  movel([0.884555, -1.427485, -2.532187, -0.752717, 1.570796, 2.455351],accel_mss,speed_ms,0,blend_radius_m)
  movel([0.882472, -1.425289, -2.533888, -0.753212, 1.570796, 2.453269],accel_mss,speed_ms,0,blend_radius_m)
  movel([0.880172, -1.423445, -2.535310, -0.753634, 1.570796, 2.450968],accel_mss,speed_ms,0,blend_radius_m)
  movel([0.877640, -1.422059, -2.536376, -0.753954, 1.570796, 2.448436],accel_mss,speed_ms,0,blend_radius_m)
  movel([0.874862, -1.421244, -2.537001, -0.754144, 1.570796, 2.445659],accel_mss,speed_ms,0,blend_radius_m)
  movel([0.871835, -1.421105, -2.537107, -0.754176, 1.570796, 2.442632],accel_mss,speed_ms,0,blend_radius_m)
  movel([0.870223, -1.421323, -2.536941, -0.754125, 1.570796, 2.441020],accel_mss,speed_ms,0,blend_radius_m)
  movel([0.868546, -1.421751, -2.536612, -0.754026, 1.570796, 2.439343],accel_mss,speed_ms,0,blend_radius_m)
  movel([0.866805, -1.422398, -2.536116, -0.753876, 1.570796, 2.437602],accel_mss,speed_ms,0,blend_radius_m)
  movel([0.864998, -1.423279, -2.535438, -0.753672, 1.570796, 2.435795],accel_mss,speed_ms,0,blend_radius_m)
  movel([0.863126, -1.424408, -2.534568, -0.753413, 1.570796, 2.433922],accel_mss,speed_ms,0,blend_radius_m)
  movel([0.861186, -1.425793, -2.533498, -0.753098, 1.570796, 2.431983],accel_mss,speed_ms,0,blend_radius_m)
  movel([0.857116, -1.429381, -2.530713, -0.752295, 1.570796, 2.427913],accel_mss,speed_ms,0,blend_radius_m)
  movel([0.855551, -1.431369, -2.529162, -0.751858, 1.570796, 2.426347],accel_mss,speed_ms,0,blend_radius_m)
  movel([0.854303, -1.433511, -2.527484, -0.751394, 1.570796, 2.425099],accel_mss,speed_ms,0,blend_radius_m)
  movel([0.853405, -1.435798, -2.525685, -0.750906, 1.570796, 2.424201],accel_mss,speed_ms,0,blend_radius_m)
  movel([0.852892, -1.438208, -2.523780, -0.750401, 1.570796, 2.423689],accel_mss,speed_ms,0,blend_radius_m)
  movel([0.855877, -1.436277, -2.525307, -0.750805, 1.570796, 2.426673],accel_mss,speed_ms,0,blend_radius_m)
  movel([0.858873, -1.434656, -2.526584, -0.751149, 1.570796, 2.429669],accel_mss,speed_ms,0,blend_radius_m)
  movel([0.861853, -1.433345, -2.527614, -0.751430, 1.570796, 2.432650],accel_mss,speed_ms,0,blend_radius_m)
  movel([0.864795, -1.432344, -2.528399, -0.751646, 1.570796, 2.435591],accel_mss,speed_ms,0,blend_radius_m)
  movel([0.867669, -1.431649, -2.528943, -0.751797, 1.570796, 2.438465],accel_mss,speed_ms,0,blend_radius_m)
  movel([0.870454, -1.431262, -2.529246, -0.751881, 1.570796, 2.441251],accel_mss,speed_ms,0,blend_radius_m)
  movel([0.873123, -1.431180, -2.529310, -0.751899, 1.570796, 2.443919],accel_mss,speed_ms,0,blend_radius_m)
  movel([0.875652, -1.431400, -2.529138, -0.751851, 1.570796, 2.446448],accel_mss,speed_ms,0,blend_radius_m)
  movel([0.878017, -1.431917, -2.528733, -0.751739, 1.570796, 2.448814],accel_mss,speed_ms,0,blend_radius_m)
  movel([0.880192, -1.432728, -2.528099, -0.751563, 1.570796, 2.450988],accel_mss,speed_ms,0,blend_radius_m)
  movel([0.882158, -1.433826, -2.527237, -0.751326, 1.570796, 2.452955],accel_mss,speed_ms,0,blend_radius_m)
  movel([0.883892, -1.435206, -2.526151, -0.751032, 1.570796, 2.454688],accel_mss,speed_ms,0,blend_radius_m)
  movel([0.885368, -1.436864, -2.524843, -0.750682, 1.570796, 2.456164],accel_mss,speed_ms,0,blend_radius_m)
  movel([0.886567, -1.438794, -2.523316, -0.750280, 1.570796, 2.457363],accel_mss,speed_ms,0,blend_radius_m)
  movel([0.887471, -1.440987, -2.521573, -0.749829, 1.570796, 2.458268],accel_mss,speed_ms,0,blend_radius_m)
  movel([0.888060, -1.443433, -2.519620, -0.749336, 1.570796, 2.458856],accel_mss,speed_ms,0,blend_radius_m)
  movel([0.888277, -1.445578, -2.517901, -0.748910, 1.570796, 2.459074],accel_mss,speed_ms,0,blend_radius_m)
  movel([0.888247, -1.447736, -2.516164, -0.748489, 1.570796, 2.459044],accel_mss,speed_ms,0,blend_radius_m)
  movel([0.887981, -1.449897, -2.514417, -0.748075, 1.570796, 2.458777],accel_mss,speed_ms,0,blend_radius_m)
  movel([0.887497, -1.452052, -2.512668, -0.747669, 1.570796, 2.458293],accel_mss,speed_ms,0,blend_radius_m)
  movel([0.885935, -1.456297, -2.509202, -0.746890, 1.570796, 2.456731],accel_mss,speed_ms,0,blend_radius_m)
  movel([0.883678, -1.460389, -2.505835, -0.746165, 1.570796, 2.454474],accel_mss,speed_ms,0,blend_radius_m)
  movel([0.880843, -1.464253, -2.502633, -0.745504, 1.570796, 2.451640],accel_mss,speed_ms,0,blend_radius_m)
  movel([0.877544, -1.467808, -2.499665, -0.744916, 1.570796, 2.448340],accel_mss,speed_ms,0,blend_radius_m)
  movel([0.873883, -1.470985, -2.496997, -0.744407, 1.570796, 2.444680],accel_mss,speed_ms,0,blend_radius_m)
  movel([0.869973, -1.473710, -2.494696, -0.743983, 1.570796, 2.440769],accel_mss,speed_ms,0,blend_radius_m)
  movel([0.865908, -1.475909, -2.492831, -0.743649, 1.570796, 2.436704],accel_mss,speed_ms,0,blend_radius_m)
  movel([0.861791, -1.477510, -2.491468, -0.743411, 1.570796, 2.432587],accel_mss,speed_ms,0,blend_radius_m)
  movel([0.857716, -1.478440, -2.490675, -0.743274, 1.570796, 2.428513],accel_mss,speed_ms,0,blend_radius_m)
  movel([0.855725, -1.478628, -2.490514, -0.743247, 1.570796, 2.426521],accel_mss,speed_ms,0,blend_radius_m)
  movel([0.853779, -1.478622, -2.490519, -0.743248, 1.570796, 2.424575],accel_mss,speed_ms,0,blend_radius_m)
  movel([0.851893, -1.478406, -2.490704, -0.743279, 1.570796, 2.422689],accel_mss,speed_ms,0,blend_radius_m)
  movel([0.850076, -1.477974, -2.491072, -0.743343, 1.570796, 2.420872],accel_mss,speed_ms,0,blend_radius_m)
  movel([0.848340, -1.477314, -2.491635, -0.743440, 1.570796, 2.419136],accel_mss,speed_ms,0,blend_radius_m)
  movel([0.846698, -1.476415, -2.492400, -0.743574, 1.570796, 2.417495],accel_mss,speed_ms,0,blend_radius_m)
  movel([0.845164, -1.475265, -2.493378, -0.743746, 1.570796, 2.415961],accel_mss,speed_ms,0,blend_radius_m)
  movel([0.843749, -1.473854, -2.494574, -0.743961, 1.570796, 2.414545],accel_mss,speed_ms,0,blend_radius_m)
  movel([0.842462, -1.472170, -2.495998, -0.744221, 1.570796, 2.413258],accel_mss,speed_ms,0,blend_radius_m)
  movel([0.841321, -1.470199, -2.497659, -0.744531, 1.570796, 2.412117],accel_mss,speed_ms,0,blend_radius_m)
  movel([0.840724, -1.468382, -2.499184, -0.744823, 1.570796, 2.411520],accel_mss,speed_ms,0,blend_radius_m)
  movel([0.839611, -1.463053, -2.503630, -0.745706, 1.570796, 2.410407],accel_mss,speed_ms,0,blend_radius_m)
  movel([0.839180, -1.459116, -2.506885, -0.746387, 1.570796, 2.409976],accel_mss,speed_ms,0,blend_radius_m)
  movel([0.839010, -1.454349, -2.510796, -0.747244, 1.570796, 2.409807],accel_mss,speed_ms,0,blend_radius_m)
  movel([0.839236, -1.448760, -2.515337, -0.748292, 1.570796, 2.410032],accel_mss,speed_ms,0,blend_radius_m)
  movel([0.840004, -1.442353, -2.520484, -0.749553, 1.570796, 2.410800],accel_mss,speed_ms,0,blend_radius_m)
  movel([0.840946, -1.437743, -2.524148, -0.750498, 1.570796, 2.411743],accel_mss,speed_ms,0,blend_radius_m)
  movel([0.842220, -1.433477, -2.527511, -0.751401, 1.570796, 2.413016],accel_mss,speed_ms,0,blend_radius_m)
  movel([0.843773, -1.429550, -2.530582, -0.752257, 1.570796, 2.414569],accel_mss,speed_ms,0,blend_radius_m)
  movel([0.845553, -1.425961, -2.533368, -0.753060, 1.570796, 2.416349],accel_mss,speed_ms,0,blend_radius_m)
  movel([0.847513, -1.422699, -2.535884, -0.753806, 1.570796, 2.418309],accel_mss,speed_ms,0,blend_radius_m)
  movel([0.849590, -1.419764, -2.538134, -0.754491, 1.570796, 2.420387],accel_mss,speed_ms,0,blend_radius_m)
  movel([0.851736, -1.417150, -2.540128, -0.755112, 1.570796, 2.422532],accel_mss,speed_ms,0,blend_radius_m)
  movel([0.853892, -1.414848, -2.541874, -0.755667, 1.570796, 2.424689],accel_mss,speed_ms,0,blend_radius_m)
  movel([0.858013, -1.411155, -2.544660, -0.756573, 1.570796, 2.428809],accel_mss,speed_ms,0,blend_radius_m)
